		IF fbFaultInjector.Status.xBusy THEN
			iTakeSlot := 1;
			iPutSlot := 1;
			IF fbFaultInjector.xWrongOperation THEN
				eActualOperation := E_MAGAZINE_OPERATION.NONE;
			ELSIF fbFaultInjector.xNoFreeSlot THEN
				eActualOperation := E_MAGAZINE_OPERATION.PUT;
			ELSE
				eActualOperation := E_MAGAZINE_OPERATION.TAKE;
			END_IF;
			Diag.eState := E_MAGAZINE_STATE.CHOOSE;
		ELSIF xFinishedLatched OR xFinishedCondition THEN
			Diag.eState := E_MAGAZINE_STATE.DISABLED;
		// Активный автоматический цикл сначала должен передать владение второму
		// магазину. До этого сохраняем xEnabled + xDisablePending, иначе менеджер
		// остаётся владельцем уже выключенного магазина и не может продолжить груз.
		ELSIF xDisableRequest
		AND NOT xRobotInMagazineContext THEN
			Diag.eState := E_MAGAZINE_STATE.DISABLED;
		ELSIF xGlobalError THEN
			Error.dwErrorActive := Error.dwErrorActive OR ERR_GLOBAL_STOP;
			Diag.eState := E_MAGAZINE_STATE.ERROR;
		// Автоматический владелец держит xExecute до завершения операции. Если
		// команда пришла раньше включения магазина, фронт был бы поглощён в
		// DISABLED; в IDLE принимаем также активный уровень запроса.
		ELSIF (rtExecute.Q OR xExecuteRequest) AND xMechanismReady THEN
			IF xManualCommand THEN
				CASE stHmiCommand.eSetPoint OF
					E_POINT_NAME.MAGAZINE_TAKE_DETAIL:
						eActualOperation := E_MAGAZINE_OPERATION.TAKE;
						iTakeSlot := stHmiCommand.iActiveSlot;
					E_POINT_NAME.MAGAZINE_PUT_DETAIL:
						eActualOperation := E_MAGAZINE_OPERATION.PUT;
						iPutSlot := stHmiCommand.iActiveSlot;
					E_POINT_NAME.MAGAZINE_CHANGE_DETAIL:
						// CHANGE требует двух слотов и запускается через ST_MAGAZINE_COMMAND.
						eActualOperation := E_MAGAZINE_OPERATION.NONE;
					E_POINT_NAME.MAGAZINE_RETURN_BLANK:
						eActualOperation := E_MAGAZINE_OPERATION.RETURN_BLANK;
						iPutSlot := stHmiCommand.iActiveSlot;
				ELSE
						eActualOperation := E_MAGAZINE_OPERATION.NONE;
				END_CASE;
			ELSE
				eActualOperation := stMagazineCommand.eOperation;
				iTakeSlot := stMagazineCommand.iTakeSlot;
				iPutSlot := stMagazineCommand.iPutSlot;
			END_IF;

			Diag.eState := E_MAGAZINE_STATE.CHOOSE;
		END_IF;

	E_MAGAZINE_STATE.CHOOSE:
		xTakeSlotValid := (iTakeSlot >= 1) AND (iTakeSlot <= iActiveSlotCount);
		xPutSlotValid := (iPutSlot >= 1) AND (iPutSlot <= iActiveSlotCount);
		xChangeTakeFirst := (eActualOperation = E_MAGAZINE_OPERATION.CHANGE)
			AND (iTakeSlot = iPutSlot);
		xTakeSlotHasBlank := FALSE;
		xPutSlotEmpty := FALSE;

		IF xTakeSlotValid THEN
		xTakeSlotHasBlank := stInventory.aSlots[iTakeSlot].xInPosition
			AND (stInventory.aSlots[iTakeSlot].eDetailType = E_DETAIL_TYPE.BLANK)
			AND (stInventory.aSlots[iTakeSlot].uiProductType >= UINT#1)
			AND (stInventory.aSlots[iTakeSlot].uiProductType <= uiTypeCount);
		END_IF;

	IF xPutSlotValid THEN
		xPutSlotEmpty := NOT stInventory.aSlots[iPutSlot].xInPosition;
	END_IF;
	xPutProductTypeValid := TRUE;
	IF (eActualOperation = E_MAGAZINE_OPERATION.PUT)
	OR (eActualOperation = E_MAGAZINE_OPERATION.CHANGE) THEN
		xPutProductTypeValid := (stRobotStatus.uiDetailPayloadType >= UINT#1)
			AND (stRobotStatus.uiDetailPayloadType <= uiTypeCount);
	ELSIF eActualOperation = E_MAGAZINE_OPERATION.RETURN_BLANK THEN
		xPutProductTypeValid := (stRobotStatus.uiBlankPayloadType >= UINT#1)
			AND (stRobotStatus.uiBlankPayloadType <= uiTypeCount);
	END_IF;

		IF fbFaultInjector.xGeometry
		OR (iActiveSlotCount = 0) THEN
			Error.dwErrorActive := Error.dwErrorActive OR ERR_GEOMETRY;
			Diag.eState := E_MAGAZINE_STATE.ERROR;

		ELSIF fbFaultInjector.xWrongOperation
		OR (eActualOperation = E_MAGAZINE_OPERATION.NONE) THEN
			Error.dwErrorActive := Error.dwErrorActive OR ERR_WRONG_OPERATION;
			Diag.eState := E_MAGAZINE_STATE.ERROR;

		ELSIF fbFaultInjector.xNoBlank THEN
			Error.dwErrorActive := Error.dwErrorActive OR ERR_NO_BLANK;
			Diag.eState := E_MAGAZINE_STATE.ERROR;

		ELSIF fbFaultInjector.xNoFreeSlot THEN
			Error.dwErrorActive := Error.dwErrorActive OR ERR_NO_FREE_SLOT;
			Diag.eState := E_MAGAZINE_STATE.ERROR;

		ELSIF fbFaultInjector.xInvalidSlot THEN
			Error.dwErrorActive := Error.dwErrorActive OR ERR_INVALID_SLOT;
			Diag.eState := E_MAGAZINE_STATE.ERROR;

		ELSIF fbFaultInjector.xSlotContent THEN
			Error.dwErrorActive := Error.dwErrorActive OR ERR_SLOT_CONTENT;
			Diag.eState := E_MAGAZINE_STATE.ERROR;

		ELSIF ((eActualOperation = E_MAGAZINE_OPERATION.TAKE)
			OR (eActualOperation = E_MAGAZINE_OPERATION.CHANGE))
		AND NOT xTakeSlotValid THEN
			Error.dwErrorActive := Error.dwErrorActive OR ERR_NO_BLANK OR ERR_INVALID_SLOT;
			Diag.eState := E_MAGAZINE_STATE.ERROR;

		ELSIF ((eActualOperation = E_MAGAZINE_OPERATION.PUT)
			OR (eActualOperation = E_MAGAZINE_OPERATION.CHANGE)
			OR (eActualOperation = E_MAGAZINE_OPERATION.RETURN_BLANK))
		AND NOT xPutSlotValid THEN
			Error.dwErrorActive := Error.dwErrorActive OR ERR_NO_FREE_SLOT OR ERR_INVALID_SLOT;
			Diag.eState := E_MAGAZINE_STATE.ERROR;

		ELSIF ((eActualOperation = E_MAGAZINE_OPERATION.TAKE)
			OR (eActualOperation = E_MAGAZINE_OPERATION.CHANGE))
		AND NOT xTakeSlotHasBlank THEN
			Error.dwErrorActive := Error.dwErrorActive OR ERR_SLOT_CONTENT;
			Diag.eState := E_MAGAZINE_STATE.ERROR;

		ELSIF ((eActualOperation = E_MAGAZINE_OPERATION.PUT)
			OR (eActualOperation = E_MAGAZINE_OPERATION.CHANGE)
			OR (eActualOperation = E_MAGAZINE_OPERATION.RETURN_BLANK))
		AND NOT xPutSlotEmpty
		AND NOT (xChangeTakeFirst AND xTakeSlotHasBlank) THEN
			Error.dwErrorActive := Error.dwErrorActive OR ERR_SLOT_CONTENT;
			Diag.eState := E_MAGAZINE_STATE.ERROR;

		ELSIF ((eActualOperation = E_MAGAZINE_OPERATION.PUT)
			OR (eActualOperation = E_MAGAZINE_OPERATION.CHANGE)
			OR (eActualOperation = E_MAGAZINE_OPERATION.RETURN_BLANK))
		AND NOT xPutProductTypeValid THEN
			Error.dwErrorActive := Error.dwErrorActive OR ERR_SLOT_CONTENT;
			Diag.eState := E_MAGAZINE_STATE.ERROR;

		ELSIF (eActualOperation = E_MAGAZINE_OPERATION.TAKE)
		AND (stRobotStatus.xBlankAvailable OR stRobotStatus.xDetailAvailable) THEN
			Error.dwErrorActive := Error.dwErrorActive OR ERR_WRONG_OPERATION;
			Diag.eState := E_MAGAZINE_STATE.ERROR;

		ELSIF (eActualOperation = E_MAGAZINE_OPERATION.CHANGE)
		AND (NOT stRobotStatus.xGripper1Open
			OR stRobotStatus.xBlankAvailable) THEN
			Error.dwErrorActive := Error.dwErrorActive OR ERR_WRONG_OPERATION;
			Diag.eState := E_MAGAZINE_STATE.ERROR;

		ELSIF ((eActualOperation = E_MAGAZINE_OPERATION.PUT)
			OR (eActualOperation = E_MAGAZINE_OPERATION.CHANGE))
		AND NOT stRobotStatus.xDetailAvailable THEN
			Error.dwErrorActive := Error.dwErrorActive OR ERR_WRONG_OPERATION;
			Diag.eState := E_MAGAZINE_STATE.ERROR;

		ELSIF (eActualOperation = E_MAGAZINE_OPERATION.RETURN_BLANK)
		AND (NOT stRobotStatus.xBlankAvailable
			OR stRobotStatus.xDetailAvailable) THEN
			Error.dwErrorActive := Error.dwErrorActive OR ERR_WRONG_OPERATION;
			Diag.eState := E_MAGAZINE_STATE.ERROR;

		ELSE
			uiPutProductType := UINT#0;
			IF (eActualOperation = E_MAGAZINE_OPERATION.PUT)
			OR (eActualOperation = E_MAGAZINE_OPERATION.CHANGE) THEN
				uiPutProductType := stRobotStatus.uiDetailPayloadType;
			ELSIF eActualOperation = E_MAGAZINE_OPERATION.RETURN_BLANK THEN
				uiPutProductType := stRobotStatus.uiBlankPayloadType;
			END_IF;
			xInventoryCommitted := FALSE;
			xTakeSlotCommitted := FALSE;
			xPutSlotCommitted := FALSE;
			xOperationSequenceComplete := FALSE;
			uiStep := 0;
			Diag.eState := E_MAGAZINE_STATE.PREPARE_STEP;
		END_IF;

	E_MAGAZINE_STATE.PREPARE_STEP:
		xRobotCommandStarted := FALSE;
		stActiveRobotCommand.xExecute := FALSE;
		stActiveRobotCommand.xStop := FALSE;
		stActiveRobotCommand.xReset := xResetRequest;
		stActiveRobotCommand.eAction := E_ROBOT_ACTION.NONE;
		stActiveRobotCommand.eSetPoint := E_POINT_NAME.NONE;

		CASE eActualOperation OF
			E_MAGAZINE_OPERATION.TAKE:
				iActiveSlot := iTakeSlot;
			E_MAGAZINE_OPERATION.PUT,
			E_MAGAZINE_OPERATION.RETURN_BLANK:
				iActiveSlot := iPutSlot;
			E_MAGAZINE_OPERATION.CHANGE:
				IF uiStep <= UINT#5 THEN
					iActiveSlot := iPutSlot;
				ELSE
					iActiveSlot := iTakeSlot;
				END_IF;
		ELSE
			iActiveSlot := SINT#0;
		END_CASE;
		stActiveRobotCommand.iActiveSlot := iActiveSlot;
		stActiveRobotCommand.uiMagazineId := uiMagazineId;

		CASE eActualOperation OF
				E_MAGAZINE_OPERATION.TAKE:
					CASE uiStep OF
						0:
							IF stRobotStatus.xRotatedToDetail THEN
								Diag.eState := E_MAGAZINE_STATE.NEXT;
							ELSE
								stActiveRobotCommand.eAction := E_ROBOT_ACTION.ROTATE_TO_DETAIL;
							END_IF;
						1:
							stActiveRobotCommand.eAction := E_ROBOT_ACTION.MOVE_TO_POINT;
							stActiveRobotCommand.eSetPoint := E_POINT_NAME.MAGAZINE_SAFE;
						2:
							stActiveRobotCommand.eAction := E_ROBOT_ACTION.MOVE_TO_POINT;
							stActiveRobotCommand.eSetPoint := E_POINT_NAME.MAGAZINE_IN_SLOT;
						3: stActiveRobotCommand.eAction := E_ROBOT_ACTION.CLAMP_1;
						4:
							stActiveRobotCommand.eAction := E_ROBOT_ACTION.MOVE_TO_POINT;
							stActiveRobotCommand.eSetPoint := E_POINT_NAME.MAGAZINE_SAFE;
					ELSE
						xOperationSequenceComplete := TRUE;
						Diag.eState := E_MAGAZINE_STATE.DONE;
					END_CASE;

				E_MAGAZINE_OPERATION.PUT:
					CASE uiStep OF
						0:
							IF stRobotStatus.xRotatedToBlank THEN
								Diag.eState := E_MAGAZINE_STATE.NEXT;
							ELSE
								stActiveRobotCommand.eAction := E_ROBOT_ACTION.ROTATE_TO_BLANK;
							END_IF;
						1:
							stActiveRobotCommand.eAction := E_ROBOT_ACTION.MOVE_TO_POINT;
							stActiveRobotCommand.eSetPoint := E_POINT_NAME.MAGAZINE_SAFE;
						2:
							stActiveRobotCommand.eAction := E_ROBOT_ACTION.MOVE_TO_POINT;
							stActiveRobotCommand.eSetPoint := E_POINT_NAME.MAGAZINE_IN_SLOT;
						3: stActiveRobotCommand.eAction := E_ROBOT_ACTION.UNCLAMP_2;
						4:
							stActiveRobotCommand.eAction := E_ROBOT_ACTION.MOVE_TO_POINT;
							stActiveRobotCommand.eSetPoint := E_POINT_NAME.MAGAZINE_SAFE;
					ELSE
						xOperationSequenceComplete := TRUE;
						Diag.eState := E_MAGAZINE_STATE.DONE;
					END_CASE;

				E_MAGAZINE_OPERATION.CHANGE:
					CASE uiStep OF
						0:
							IF (xChangeTakeFirst AND stRobotStatus.xRotatedToDetail)
							OR (NOT xChangeTakeFirst AND stRobotStatus.xRotatedToBlank) THEN
								Diag.eState := E_MAGAZINE_STATE.NEXT;
							ELSIF xChangeTakeFirst THEN
								stActiveRobotCommand.eAction := E_ROBOT_ACTION.ROTATE_TO_DETAIL;
							ELSE
								stActiveRobotCommand.eAction := E_ROBOT_ACTION.ROTATE_TO_BLANK;
							END_IF;
						1:
							stActiveRobotCommand.eAction := E_ROBOT_ACTION.MOVE_TO_POINT;
							stActiveRobotCommand.eSetPoint := E_POINT_NAME.MAGAZINE_SAFE;
						2:
							stActiveRobotCommand.eAction := E_ROBOT_ACTION.MOVE_TO_POINT;
							stActiveRobotCommand.eSetPoint := E_POINT_NAME.MAGAZINE_IN_SLOT;
						3:
							IF xChangeTakeFirst THEN
								stActiveRobotCommand.eAction := E_ROBOT_ACTION.CLAMP_1;
							ELSE
								stActiveRobotCommand.eAction := E_ROBOT_ACTION.UNCLAMP_2;
							END_IF;
						4:
							stActiveRobotCommand.eAction := E_ROBOT_ACTION.MOVE_TO_POINT;
							stActiveRobotCommand.eSetPoint := E_POINT_NAME.MAGAZINE_CHANGE;
						5:
							IF (xChangeTakeFirst AND stRobotStatus.xRotatedToBlank)
							OR (NOT xChangeTakeFirst AND stRobotStatus.xRotatedToDetail) THEN
								Diag.eState := E_MAGAZINE_STATE.NEXT;
							ELSIF xChangeTakeFirst THEN
								stActiveRobotCommand.eAction := E_ROBOT_ACTION.ROTATE_TO_BLANK;
							ELSE
								stActiveRobotCommand.eAction := E_ROBOT_ACTION.ROTATE_TO_DETAIL;
							END_IF;
						6:
							stActiveRobotCommand.eAction := E_ROBOT_ACTION.MOVE_TO_POINT;
							stActiveRobotCommand.eSetPoint := E_POINT_NAME.MAGAZINE_CHANGE;
						7:
							stActiveRobotCommand.eAction := E_ROBOT_ACTION.MOVE_TO_POINT;
							stActiveRobotCommand.eSetPoint := E_POINT_NAME.MAGAZINE_IN_SLOT;
						8:
							IF xChangeTakeFirst THEN
								stActiveRobotCommand.eAction := E_ROBOT_ACTION.UNCLAMP_2;
							ELSE
								stActiveRobotCommand.eAction := E_ROBOT_ACTION.CLAMP_1;
							END_IF;
						9:
							stActiveRobotCommand.eAction := E_ROBOT_ACTION.MOVE_TO_POINT;
							stActiveRobotCommand.eSetPoint := E_POINT_NAME.MAGAZINE_SAFE;
					ELSE
						xOperationSequenceComplete := TRUE;
						Diag.eState := E_MAGAZINE_STATE.DONE;
					END_CASE;

				E_MAGAZINE_OPERATION.RETURN_BLANK:
					CASE uiStep OF
						0:
							IF stRobotStatus.xRotatedToDetail THEN
								Diag.eState := E_MAGAZINE_STATE.NEXT;
							ELSE
								stActiveRobotCommand.eAction := E_ROBOT_ACTION.ROTATE_TO_DETAIL;
							END_IF;
						1:
							stActiveRobotCommand.eAction := E_ROBOT_ACTION.MOVE_TO_POINT;
							stActiveRobotCommand.eSetPoint := E_POINT_NAME.MAGAZINE_SAFE;
						2:
							stActiveRobotCommand.eAction := E_ROBOT_ACTION.MOVE_TO_POINT;
							stActiveRobotCommand.eSetPoint := E_POINT_NAME.MAGAZINE_IN_SLOT;
						3: stActiveRobotCommand.eAction := E_ROBOT_ACTION.UNCLAMP_1;
						4:
							stActiveRobotCommand.eAction := E_ROBOT_ACTION.MOVE_TO_POINT;
							stActiveRobotCommand.eSetPoint := E_POINT_NAME.MAGAZINE_SAFE;
					ELSE
						xOperationSequenceComplete := TRUE;
						Diag.eState := E_MAGAZINE_STATE.DONE;
					END_CASE;
		END_CASE;

		IF Diag.eState = E_MAGAZINE_STATE.PREPARE_STEP THEN
			Diag.eState := E_MAGAZINE_STATE.ROBOT_COMMAND;
		END_IF;

	E_MAGAZINE_STATE.ROBOT_COMMAND:
		Command := stActiveRobotCommand;
		Command.xExecute := TRUE;
		IF stRobotStatus.xBusy THEN
			xRobotCommandStarted := TRUE;
		END_IF;

		IF xStopRequest OR xGlobalError THEN
			Command.xStop := stRobotStatus.xBusy;
			Error.dwErrorActive := Error.dwErrorActive OR ERR_GLOBAL_STOP;
			Diag.eState := E_MAGAZINE_STATE.ERROR;

		ELSIF stRobotStatus.xError THEN
			Error.dwErrorActive := Error.dwErrorActive OR ERR_ROBOT;
			Diag.eState := E_MAGAZINE_STATE.ERROR;

		ELSIF xRobotCommandStarted AND stRobotStatus.xDone THEN
			// Матрица меняется в момент подтверждённого физического переноса,
			// а не после отхода робота и завершения всей составной операции.
			CASE eActualOperation OF
				E_MAGAZINE_OPERATION.TAKE:
					IF (uiStep = UINT#3) AND NOT xTakeSlotCommitted THEN
						stInventory.aSlots[iTakeSlot].xInPosition := FALSE;
						stInventory.aSlots[iTakeSlot].eDetailType := E_DETAIL_TYPE.NONE;
						stInventory.aSlots[iTakeSlot].uiProductType := UINT#0;
						xTakeSlotCommitted := TRUE;
					END_IF;

				E_MAGAZINE_OPERATION.PUT:
					IF (uiStep = UINT#3) AND NOT xPutSlotCommitted THEN
						stInventory.aSlots[iPutSlot].xInPosition := TRUE;
						stInventory.aSlots[iPutSlot].eDetailType := E_DETAIL_TYPE.DETAIL;
						stInventory.aSlots[iPutSlot].uiProductType := uiPutProductType;
						udiProducedPartsTotal := udiProducedPartsTotal + UDINT#1;
						xPutSlotCommitted := TRUE;
					END_IF;

				E_MAGAZINE_OPERATION.CHANGE:
					IF (((uiStep = UINT#3) AND NOT xChangeTakeFirst)
						OR ((uiStep = UINT#8) AND xChangeTakeFirst))
					AND NOT xPutSlotCommitted THEN
						stInventory.aSlots[iPutSlot].xInPosition := TRUE;
						stInventory.aSlots[iPutSlot].eDetailType := E_DETAIL_TYPE.DETAIL;
						stInventory.aSlots[iPutSlot].uiProductType := uiPutProductType;
						udiProducedPartsTotal := udiProducedPartsTotal + UDINT#1;
						xPutSlotCommitted := TRUE;
					ELSIF (((uiStep = UINT#8) AND NOT xChangeTakeFirst)
						OR ((uiStep = UINT#3) AND xChangeTakeFirst))
					AND NOT xTakeSlotCommitted THEN
						stInventory.aSlots[iTakeSlot].xInPosition := FALSE;
						stInventory.aSlots[iTakeSlot].eDetailType := E_DETAIL_TYPE.NONE;
						stInventory.aSlots[iTakeSlot].uiProductType := UINT#0;
						xTakeSlotCommitted := TRUE;
					END_IF;

				E_MAGAZINE_OPERATION.RETURN_BLANK:
					IF (uiStep = UINT#3) AND NOT xPutSlotCommitted THEN
						xFinishedLatched := FALSE;
						xFinishedCondition := FALSE;
						stInventory.aSlots[iPutSlot].xInPosition := TRUE;
						stInventory.aSlots[iPutSlot].eDetailType := E_DETAIL_TYPE.BLANK;
						stInventory.aSlots[iPutSlot].uiProductType := uiPutProductType;
						xPutSlotCommitted := TRUE;
					END_IF;
			END_CASE;
			Diag.eState := E_MAGAZINE_STATE.RELEASE_ROBOT_COMMAND;
		END_IF;

	E_MAGAZINE_STATE.RELEASE_ROBOT_COMMAND:
		IF stRobotStatus.xError THEN
			Error.dwErrorActive := Error.dwErrorActive OR ERR_ROBOT;
			Diag.eState := E_MAGAZINE_STATE.ERROR;
		ELSIF NOT stRobotStatus.xBusy AND NOT stRobotStatus.xDone THEN
			Diag.eState := E_MAGAZINE_STATE.NEXT;
		END_IF;

	E_MAGAZINE_STATE.NEXT:
		uiStep := uiStep + 1;
		Diag.eState := E_MAGAZINE_STATE.PREPARE_STEP;

	E_MAGAZINE_STATE.DONE:
		// Страховочная фиксация нужна только если конечный DONE получен без
		// промежуточного обновления. В штатном ходе слоты уже изменены захватами.
		IF xOperationSequenceComplete
		AND NOT xStopRequest
		AND NOT xGlobalError
		AND NOT xInventoryCommitted THEN
			CASE eActualOperation OF
				E_MAGAZINE_OPERATION.TAKE:
					IF NOT xTakeSlotCommitted THEN
						stInventory.aSlots[iTakeSlot].xInPosition := FALSE;
						stInventory.aSlots[iTakeSlot].eDetailType := E_DETAIL_TYPE.NONE;
						stInventory.aSlots[iTakeSlot].uiProductType := UINT#0;
						xTakeSlotCommitted := TRUE;
					END_IF;
				E_MAGAZINE_OPERATION.PUT:
					IF NOT xPutSlotCommitted THEN
						stInventory.aSlots[iPutSlot].xInPosition := TRUE;
						stInventory.aSlots[iPutSlot].eDetailType := E_DETAIL_TYPE.DETAIL;
						stInventory.aSlots[iPutSlot].uiProductType := uiPutProductType;
						udiProducedPartsTotal := udiProducedPartsTotal + UDINT#1;
						xPutSlotCommitted := TRUE;
					END_IF;
				E_MAGAZINE_OPERATION.CHANGE:
					// Для обмена в одном слоте сначала отражаем изъятие. Уже
					// подтверждённую укладку нельзя затереть страховочной фиксацией.
					IF NOT xTakeSlotCommitted THEN
						IF NOT xChangeTakeFirst OR NOT xPutSlotCommitted THEN
							stInventory.aSlots[iTakeSlot].xInPosition := FALSE;
							stInventory.aSlots[iTakeSlot].eDetailType := E_DETAIL_TYPE.NONE;
							stInventory.aSlots[iTakeSlot].uiProductType := UINT#0;
						END_IF;
						xTakeSlotCommitted := TRUE;
					END_IF;
					IF NOT xPutSlotCommitted THEN
						stInventory.aSlots[iPutSlot].xInPosition := TRUE;
						stInventory.aSlots[iPutSlot].eDetailType := E_DETAIL_TYPE.DETAIL;
						stInventory.aSlots[iPutSlot].uiProductType := uiPutProductType;
						udiProducedPartsTotal := udiProducedPartsTotal + UDINT#1;
						xPutSlotCommitted := TRUE;
					END_IF;
				E_MAGAZINE_OPERATION.RETURN_BLANK:
					IF NOT xPutSlotCommitted THEN
						xFinishedLatched := FALSE;
						xFinishedCondition := FALSE;
						stInventory.aSlots[iPutSlot].xInPosition := TRUE;
						stInventory.aSlots[iPutSlot].eDetailType := E_DETAIL_TYPE.BLANK;
						stInventory.aSlots[iPutSlot].uiProductType := uiPutProductType;
						xPutSlotCommitted := TRUE;
					END_IF;
			END_CASE;
			xInventoryCommitted := TRUE;
		END_IF;
		IF NOT xExecuteRequest THEN
			eActualOperation := E_MAGAZINE_OPERATION.NONE;
			IF xDisableRequest
			AND NOT xRobotInMagazineContext THEN
				Diag.eState := E_MAGAZINE_STATE.DISABLED;
			ELSE
				Diag.eState := E_MAGAZINE_STATE.IDLE;
			END_IF;
		END_IF;

	E_MAGAZINE_STATE.ERROR:
		IF xResetRequest
		AND NOT xIoManual
		AND NOT xExecuteRequest
		AND NOT xStopRequest
		AND NOT FaultStatus.xBusy
		AND NOT xGlobalError
		AND xRobotResetDependencyReady THEN
			Error.dwErrorLast := Error.dwErrorActive;
			Error.dwErrorActive := DWORD#0;
			eActualOperation := E_MAGAZINE_OPERATION.NONE;
			Diag.eState := E_MAGAZINE_STATE.DISABLED;
		END_IF;
END_CASE;

// Класс реакции не размазывается по CASE. Первичная причина остаётся в своей
// маске, а контекст конкретного магазина хранится до принятого сброса.
IF (Diag.eState = E_MAGAZINE_STATE.ERROR)
AND NOT xFaultContextCaptured THEN
	xRobotInMagazineAtFault := xRobotInMagazineContext;
	xFaultContextCaptured := TRUE;
ELSIF Diag.eState <> E_MAGAZINE_STATE.ERROR THEN
	xRobotInMagazineAtFault := FALSE;
	xFaultContextCaptured := FALSE;
END_IF;

xRobotStopRequired := NOT xGlobalError
	AND (
		((Error.dwErrorActive AND ERR_ROBOT) <> DWORD#0)
		OR (((Error.dwErrorActive AND MASK_EQUIPMENT_ERROR) <> DWORD#0)
			AND xRobotInMagazineAtFault)
	);

// Физический Stop нужен только занятому роботу. При неподвижном роботе внутри
// магазина FB_ROBOT получит зависимую ошибку без пустой команды остановки.
IF (Diag.eState = E_MAGAZINE_STATE.ERROR)
AND xRobotStopRequired
AND stRobotStatus.xBusy THEN
	Command := stActiveRobotCommand;
	Command.xExecute := TRUE;
	Command.xStop := TRUE;
END_IF;

// ERROR технологически отключает магазин немедленно, но причина остаётся
// защёлкнутой до разрешённого Reset.
Status.xEnabled := (Diag.eState <> E_MAGAZINE_STATE.DISABLED)
	AND (Diag.eState <> E_MAGAZINE_STATE.ERROR);
Status.xDisablePending := xDisableRequest AND Status.xEnabled;
Status.xPowerAllowed := Status.xEnabled OR Status.xEnableSequenceAllowed;
Status.xFillAllowed := (iActiveSlotCount > SINT#0) AND Status.xEditAllowed;
Status.xClearAllowed := Status.xEditAllowed;
Status.xReady := xMechanismReady AND  (Diag.eState = E_MAGAZINE_STATE.IDLE)
	AND xRobotCanWorkWithMagazine
	AND (Error.dwErrorActive = DWORD#0);
Status.xBusy := (Diag.eState <> E_MAGAZINE_STATE.DISABLED)
	AND (Diag.eState <> E_MAGAZINE_STATE.IDLE)
	AND (Diag.eState <> E_MAGAZINE_STATE.DONE)
	AND (Diag.eState <> E_MAGAZINE_STATE.ERROR);
Status.xDone := Diag.eState = E_MAGAZINE_STATE.DONE;
Status.xError := Diag.eState = E_MAGAZINE_STATE.ERROR;
Status.xRobotStopRequired := xRobotStopRequired;
Status.udiProducedPartsTotal := udiProducedPartsTotal;
Status.uiMagazineId := uiMagazineId;
Status.eGrantedOperation := eGrantedOperation;
Status.eActualOperation := eActualOperation;
Status.iSelectedBlank := iTakeSlot;
Status.iSelectedFreeSlot := iPutSlot;
// Разовая доработка палеты завершена: чужой груз/станок не возвращает её
// в планирование. Защёлку снимает только смена банка или правка его содержимого.
xFinishedLatched := xFinishedLatched OR (xFinishedCondition AND NOT Status.xBusy);
Status.xFinished := xFinishedLatched;
Error.dwAlarmActive := Error.dwErrorActive;

IF Error.dwErrorActive <> DWORD#0 THEN
	Error.dwErrorLast := Error.dwErrorActive;
END_IF;

Error.stErrorActive := UpdateErrorView(dwError := Error.dwErrorActive);
Error.stErrorLast := UpdateErrorView(dwError := Error.dwErrorLast);
FaultStatus.xResetAllowed := Status.xError
	AND NOT xIoManual
	AND NOT FaultStatus.xBusy
	AND NOT xExecuteRequest
	AND NOT xStopRequest
	AND NOT xGlobalError
	AND xRobotResetDependencyReady;

// Сводка публикуется владельцем содержимого после всех изменений слотов.
UpdateTypeStatus(stMagazineInventory := stInventory);

METHOD FindBlank : SINT
VAR_INPUT
	iSlotCount : SINT; // Число слотов, участвующих в поиске
END_VAR
VAR_IN_OUT
	stDetail : ARRAY [1..GVL_CELL_SETTINGS.NumberDetail] OF ST_DETAIL; // Содержимое слотов магазина
END_VAR
VAR
	i : SINT; // Индекс проверяемого слота
END_VAR
FindBlank := 0;

FOR i:= 1 TO iSlotCount DO
	IF stDetail[i].xInPosition = TRUE AND stDetail[i].eDetailType =  E_DETAIL_TYPE.BLANK THEN
		FindBlank := i;
		EXIT;
	END_IF
END_FOR
END_METHOD

METHOD UpdateErrorView : ST_MAGAZINE_ERROR
VAR_INPUT
	dwError : DWORD; // Битовая маска для расшифровки
END_VAR
VAR
	stError : ST_MAGAZINE_ERROR; // Представление ошибок отдельными флагами
END_VAR
stError.WRONG_OPERATION := (dwError AND ERR_WRONG_OPERATION) <> DWORD#0;
stError.NO_BLANK := (dwError AND ERR_NO_BLANK) <> DWORD#0;
stError.NO_FREE_SLOT := (dwError AND ERR_NO_FREE_SLOT) <> DWORD#0;
stError.INVALID_SLOT := (dwError AND ERR_INVALID_SLOT) <> DWORD#0;
stError.SLOT_CONTENT := (dwError AND ERR_SLOT_CONTENT) <> DWORD#0;
stError.ROBOT_ERROR := (dwError AND ERR_ROBOT) <> DWORD#0;
stError.GLOBAL_STOP := (dwError AND ERR_GLOBAL_STOP) <> DWORD#0;
stError.GEOMETRY_ERROR := (dwError AND ERR_GEOMETRY) <> DWORD#0;

UpdateErrorView := stError;
END_METHOD

METHOD FindFreeSlot : SINT
VAR_INPUT
	iSlotCount : SINT; // Число слотов, участвующих в поиске
END_VAR
VAR_IN_OUT
	stDetail : ARRAY [1..GVL_CELL_SETTINGS.NumberDetail] OF ST_DETAIL; // Содержимое слотов магазина
END_VAR
VAR
	i : SINT; // Индекс проверяемого слота
END_VAR
FindFreeSlot := 0;

FOR i:= 1 TO iSlotCount DO
	IF stDetail[i].xInPosition = FALSE THEN
		FindFreeSlot := i;
		EXIT;
	END_IF
END_FOR
END_METHOD

METHOD PRIVATE UpdateTypeStatus
VAR_IN_OUT
	stMagazineInventory : ST_MAGAZINE_INVENTORY;
END_VAR
VAR
	uiType : UINT; // Тип секции, 1..3
	uiSlot : UINT; // Проверяемый слот
	iSlot  : SINT; // Индекс массива содержимого
END_VAR
FOR uiType := UINT#1 TO UINT#3 DO
	Status.stTypeStatus.aiBlankSlot[uiType] := SINT#0;
	Status.stTypeStatus.aiFreeSlot[uiType] := SINT#0;
	Status.stTypeStatus.auiBlankCount[uiType] := UINT#0;
	Status.stTypeStatus.auiDetailCount[uiType] := UINT#0;
	Status.stTypeStatus.auiFreeCount[uiType] := UINT#0;
END_FOR;

IF (iActiveSlotCount > SINT#0)
AND (uiTypeCount >= UINT#1)
AND (uiTypeCount <= UINT#3) THEN
	FOR uiSlot := UINT#1 TO SINT_TO_UINT(iActiveSlotCount) DO
		iSlot := UINT_TO_SINT(uiSlot);
		IF NOT stMagazineInventory.aSlots[iSlot].xInPosition THEN
			// Пустой слот универсален: тип 0
			// означает отсутствие изделия, а не запрет укладки конкретного типа.
			FOR uiType := UINT#1 TO uiTypeCount DO
				Status.stTypeStatus.auiFreeCount[uiType] :=
					Status.stTypeStatus.auiFreeCount[uiType] + UINT#1;
				IF Status.stTypeStatus.aiFreeSlot[uiType] = SINT#0 THEN
					Status.stTypeStatus.aiFreeSlot[uiType] := iSlot;
				END_IF;
			END_FOR;
		ELSE
			uiType := stMagazineInventory.aSlots[iSlot].uiProductType;
			IF (uiType >= UINT#1) AND (uiType <= uiTypeCount)
			AND (stMagazineInventory.aSlots[iSlot].eDetailType = E_DETAIL_TYPE.BLANK) THEN
				Status.stTypeStatus.auiBlankCount[uiType] :=
					Status.stTypeStatus.auiBlankCount[uiType] + UINT#1;
				IF Status.stTypeStatus.aiBlankSlot[uiType] = SINT#0 THEN
					Status.stTypeStatus.aiBlankSlot[uiType] := iSlot;
				END_IF;
			ELSIF (uiType >= UINT#1) AND (uiType <= uiTypeCount)
			AND (stMagazineInventory.aSlots[iSlot].eDetailType = E_DETAIL_TYPE.DETAIL) THEN
				Status.stTypeStatus.auiDetailCount[uiType] :=
					Status.stTypeStatus.auiDetailCount[uiType] + UINT#1;
			END_IF;
		END_IF;
	END_FOR;
END_IF;
END_METHOD

END_FUNCTION_BLOCK

// Device/Application/FB/FB_FAULT_INJECTOR/FB_MAGAZINE_FAULT_INJECTOR
FUNCTION_BLOCK FB_MAGAZINE_FAULT_INJECTOR
VAR_INPUT
	Request       : ST_MAGAZINE_FAULT_REQUEST; // Запросы конкретных ошибок магазина
	xOwnerAllowed : BOOL; // Безопасные условия, рассчитанные FB_MAGAZINE
	xComplete     : BOOL; // Штатная ошибка уже сформирована владельцем
END_VAR
VAR_OUTPUT
	xWrongOperation : BOOL;
	xNoBlank        : BOOL;
	xNoFreeSlot     : BOOL;
	xInvalidSlot    : BOOL;
	xSlotContent    : BOOL;
	xGeometry       : BOOL;
	Status          : ST_FAULT_INJECTION_STATUS; // Состояние источника для HMI
END_VAR
VAR
	rtWrongOperation : R_TRIG;
	rtNoBlank        : R_TRIG;
	rtNoFreeSlot     : R_TRIG;
	rtInvalidSlot    : R_TRIG;
	rtSlotContent    : R_TRIG;
	rtGeometry       : R_TRIG;
	xRequestPulse    : BOOL;
END_VAR

rtWrongOperation(CLK := Request.xWrongOperation);
rtNoBlank(CLK := Request.xNoBlank);
rtNoFreeSlot(CLK := Request.xNoFreeSlot);
rtInvalidSlot(CLK := Request.xInvalidSlot);
rtSlotContent(CLK := Request.xSlotContent);
rtGeometry(CLK := Request.xGeometry);

xRequestPulse := rtWrongOperation.Q
	OR rtNoBlank.Q
	OR rtNoFreeSlot.Q
	OR rtInvalidSlot.Q
	OR rtSlotContent.Q
	OR rtGeometry.Q;

Status.xRejected := FALSE;
Status.xAllowed := Request.xEnabled AND xOwnerAllowed;

IF xComplete THEN
	xWrongOperation := FALSE;
	xNoBlank := FALSE;
	xNoFreeSlot := FALSE;
	xInvalidSlot := FALSE;
	xSlotContent := FALSE;
	xGeometry := FALSE;
END_IF;

IF xRequestPulse THEN
	IF Status.xAllowed THEN
		xWrongOperation := rtWrongOperation.Q;
		xNoBlank := rtNoBlank.Q;
		xNoFreeSlot := rtNoFreeSlot.Q;
		xInvalidSlot := rtInvalidSlot.Q;
		xSlotContent := rtSlotContent.Q;
		xGeometry := rtGeometry.Q;
	ELSE
		Status.xRejected := TRUE;
		Status.udiRejectSequence := Status.udiRejectSequence + UDINT#1;
		IF Status.udiRejectSequence = UDINT#0 THEN
			Status.udiRejectSequence := UDINT#1;
		END_IF;
	END_IF;
END_IF;

Status.xActive := xWrongOperation
	OR xNoBlank
	OR xNoFreeSlot
	OR xInvalidSlot
	OR xSlotContent
	OR xGeometry;
Status.xBusy := Status.xActive;
Status.xResetAllowed := FALSE;

END_FUNCTION_BLOCK

// Device/Application/FB/FB_ROBOT_MODBUS
{attribute 'no_assign'}
FUNCTION_BLOCK FB_ROBOT_MODBUS
VAR_INPUT
	xEnable          : BOOL; // Применён режим MODBUS_TCP
	xReconnect       : BOOL; // Настройки изменены, выполнить reconnect
	Config           : ST_ROBOT_MODBUS_CONFIG;
	Command          : ST_ROBOT_COMMAND; // Семантическая команда FB_ROBOT
END_VAR
VAR_OUTPUT
	Status           : ST_ROBOT_MODBUS_STATUS;
END_VAR
VAR_IN_OUT
	auiWriteRegisters : ARRAY [0..8] OF UINT; // Документные адреса 1001..1009
	auiReadRegisters  : ARRAY [0..16] OF UINT; // Документные адреса 1101..1117
END_VAR
VAR
	{attribute 'no_assign'}
	fbClient       : ModbusFB.ClientTCP;
	fbRead         : ModbusFB.ClientRequestReadHoldingRegisters;
	fbWrite        : ModbusFB.ClientRequestWriteMultipleRegisters;
	eState         : E_ROBOT_MODBUS_CLIENT_STATE := E_ROBOT_MODBUS_CLIENT_STATE.DISABLED;
	xConnect       : BOOL;
	xReadExecute   : BOOL;
	xWriteExecute  : BOOL;
	xStatusFresh   : BOOL;
	xCommandArmed  : BOOL;
	xCommandActive : BOOL;
	xWritePending  : BOOL;
	xHeartbeatChanged : BOOL;
	xHeartbeatSeen : BOOL;
	xPlcHeartbeatDue : BOOL;
	xStopPending   : BOOL;
	xResetPending  : BOOL;
	xResetInProgress : BOOL;
	xResetWriteDone : BOOL; // FC16 с Reset=1 подтверждена сервером
	tonResetAttempt : TON;
	xControlClearPending : BOOL;
	rtStop         : R_TRIG;
	rtReset        : R_TRIG;
	rtReconnect    : R_TRIG;
	tonPoll        : TON;
	tonPlcHeartbeat: TON;
	tonRobotHeartbeat : TON;
	tonCommunicationGrace : TON;
	tonCommandTimeout : TON;
	tonReconnect   : TON;
	uiCommandSeq   : UINT;
	uiActiveSeq    : UINT;
	uiDecodedRobotHeartbeat : UINT; // Heartbeat из последнего завершённого FC03
	uiPositionXHigh : UINT; // Координаты из того же завершённого FC03-снимка
	uiPositionXLow  : UINT;
	uiPositionYHigh : UINT;
	uiPositionYLow  : UINT;
	uiPositionZHigh : UINT;
	uiPositionZLow  : UINT;
	uiPlcHeartbeat : UINT;
	uiLastRobotHeartbeat : UINT;
	uiCommandCode  : UINT;
	uiRegisterIndex : UINT;
	dwPositionRaw  : DWORD;
	diPositionRaw  : DINT;
	udiReplyTimeoutUs : UDINT;
END_VAR
VAR CONSTANT
	COMMAND_START_ITEM : UINT := UINT#1000; // Документный 1001
	STATUS_START_ITEM  : UINT := UINT#1100; // Документный 1101
	COMMAND_QUANTITY   : UINT := UINT#9;
	STATUS_QUANTITY    : UINT := UINT#17;
	PROTOCOL_VERSION   : UINT := UINT#3;
	RESET_ATTEMPT_TIMEOUT : TIME := T#10S; // Полная попытка: запись, feedback, снятие
	STATUS_CONTROLLER_ON  : UINT := UINT#16#0001;
	STATUS_AUTOMATIC_MODE : UINT := UINT#16#0002;
	STATUS_REMOTE_ENABLED : UINT := UINT#16#0004;
	STATUS_DRIVES_ENABLED : UINT := UINT#16#0008;
	STATUS_HOMED          : UINT := UINT#16#0010;
	STATUS_EMERGENCY_STOP : UINT := UINT#16#0020;
	STATUS_ROBOT_ALARM    : UINT := UINT#16#0040;
	STATUS_ROBOT_READY    : UINT := UINT#16#0080;
	STATUS_POSITION_VALID : UINT := UINT#16#0100;
	STATUS_SIMULATOR_ACTIVE : UINT := UINT#16#0200;
END_VAR

Status.xConfigValid := (Config.aIpAddress[0] > BYTE#0)
	AND (Config.aIpAddress[0] < BYTE#224)
	AND (Config.uiPort > UINT#0)
	AND (Config.uiUnitId <= UINT#255)
	AND (Config.tResponseTimeout >= T#50MS)
	AND (Config.tPollInterval >= T#10MS)
	AND (Config.tHeartbeatTimeout >= T#500MS)
	AND (Config.tCommandTimeout >= T#1S);

	udiReplyTimeoutUs := TIME_TO_UDINT(Config.tResponseTimeout) * UDINT#1000;
	rtStop(CLK := Command.xStop);
	rtReset(CLK := Command.xReset);
	rtReconnect(CLK := xReconnect);
	IF rtStop.Q THEN
		xStopPending := TRUE;
	END_IF;
	IF rtReset.Q AND NOT xResetInProgress THEN
		xResetPending := TRUE;
		xResetInProgress := TRUE;
		xResetWriteDone := FALSE;
		Status.xResetDone := FALSE;
		Status.xResetFailed := FALSE;
	END_IF;
xReadExecute := FALSE;
xWriteExecute := FALSE;
xHeartbeatChanged := FALSE;

fbClient(
	xConnect := xConnect,
	aIPaddr := Config.aIpAddress,
	uiPort := Config.uiPort,
	tConnnectTimeOut := Config.tHeartbeatTimeout
);

IF NOT xEnable OR NOT Status.xConfigValid THEN
	xConnect := FALSE;
	eState := E_ROBOT_MODBUS_CLIENT_STATE.DISABLED;
	xStatusFresh := FALSE;
	xCommandArmed := FALSE;
	xCommandActive := FALSE;
	xWritePending := FALSE;
	xStopPending := FALSE;
	xResetPending := FALSE;
	xResetInProgress := FALSE;
	xResetWriteDone := FALSE;
	Status.xResetDone := FALSE;
	Status.xResetFailed := FALSE;
	xControlClearPending := FALSE;
	xHeartbeatSeen := FALSE;
	xPlcHeartbeatDue := FALSE;
	uiActiveSeq := UINT#0;
	Status.xConnected := FALSE;
ELSE
	xConnect := TRUE;
	IF rtReconnect.Q THEN
		xConnect := FALSE;
		eState := E_ROBOT_MODBUS_CLIENT_STATE.RECONNECT_WAIT;
		xStatusFresh := FALSE;
		xCommandArmed := FALSE;
		xCommandActive := FALSE;
		xWritePending := FALSE;
		xControlClearPending := FALSE;
		xHeartbeatSeen := FALSE;
		xPlcHeartbeatDue := FALSE;
	END_IF;
END_IF;

CASE eState OF
	E_ROBOT_MODBUS_CLIENT_STATE.DISABLED:
		IF xEnable AND Status.xConfigValid THEN
			xConnect := TRUE;
			eState := E_ROBOT_MODBUS_CLIENT_STATE.CONNECTING;
		END_IF;

	E_ROBOT_MODBUS_CLIENT_STATE.CONNECTING:
		IF fbClient.xConnected THEN
			eState := E_ROBOT_MODBUS_CLIENT_STATE.INITIAL_READ;
		ELSIF fbClient.xError THEN
			Status.udiClientError := TO_UDINT(fbClient.eErrorID);
			xConnect := FALSE;
			eState := E_ROBOT_MODBUS_CLIENT_STATE.RECONNECT_WAIT;
		END_IF;

	E_ROBOT_MODBUS_CLIENT_STATE.INITIAL_READ:
		xReadExecute := TRUE;
		IF fbRead.xDone THEN
			xStatusFresh := TRUE;
			uiCommandSeq := auiReadRegisters[0];
			uiActiveSeq := UINT#0;
			uiPlcHeartbeat := UINT#0;
			uiLastRobotHeartbeat := auiReadRegisters[6];
			xHeartbeatSeen := FALSE;
			FOR uiRegisterIndex := UINT#0 TO UINT#8 DO
				auiWriteRegisters[uiRegisterIndex] := UINT#0;
			END_FOR;
			auiWriteRegisters[7] := uiCommandSeq;
			eState := E_ROBOT_MODBUS_CLIENT_STATE.INITIAL_READ_RELEASE;
		ELSIF fbRead.xError THEN
			Status.udiReadError := TO_UDINT(fbRead.eErrorID);
			xConnect := FALSE;
			eState := E_ROBOT_MODBUS_CLIENT_STATE.RECONNECT_WAIT;
		END_IF;

	E_ROBOT_MODBUS_CLIENT_STATE.INITIAL_READ_RELEASE:
		IF NOT fbRead.xBusy THEN
			eState := E_ROBOT_MODBUS_CLIENT_STATE.CLEAR_COMMAND;
		END_IF;

	E_ROBOT_MODBUS_CLIENT_STATE.CLEAR_COMMAND:
		xWriteExecute := TRUE;
		IF fbWrite.xDone THEN
			eState := E_ROBOT_MODBUS_CLIENT_STATE.CLEAR_COMMAND_RELEASE;
		ELSIF fbWrite.xError THEN
			Status.udiWriteError := TO_UDINT(fbWrite.eErrorID);
			xConnect := FALSE;
			eState := E_ROBOT_MODBUS_CLIENT_STATE.RECONNECT_WAIT;
		END_IF;

	E_ROBOT_MODBUS_CLIENT_STATE.CLEAR_COMMAND_RELEASE:
		IF NOT fbWrite.xBusy THEN
			xCommandArmed := NOT Command.xExecute;
			xCommandActive := FALSE;
			eState := E_ROBOT_MODBUS_CLIENT_STATE.READY;
		END_IF;

	E_ROBOT_MODBUS_CLIENT_STATE.READY:
		IF NOT fbClient.xConnected OR fbClient.xError THEN
			Status.udiClientError := TO_UDINT(fbClient.eErrorID);
			xConnect := FALSE;
			eState := E_ROBOT_MODBUS_CLIENT_STATE.RECONNECT_WAIT;
		ELSIF xStopPending THEN
			// Stop отменяет текущую попытку сброса; он не может быть проглочен Reset.
			IF xResetInProgress THEN Status.xResetFailed := TRUE; END_IF;
			xResetInProgress := FALSE;
			xResetWriteDone := FALSE;
			// Stop always preempts Reset and normal commands.
			// Execute снимается сразу: после принятого CommandSeq это не отменяет
			// команду, зато позволяет роботу выйти из DONE/ERROR/STOPPED в IDLE.
			// Без этого уже завершённая дискретная команда навечно удерживала
			// Execute=1, а xControlClearPending ждал недостижимый IDLE.
			auiWriteRegisters[0] := UINT#0;
			auiWriteRegisters[1] := UINT#0;
			auiWriteRegisters[2] := UINT#1;
			auiWriteRegisters[3] := UINT#0;
			auiWriteRegisters[4] := UINT#0;
			auiWriteRegisters[5] := UINT#0;
			auiWriteRegisters[6] := UINT#0;
			xStopPending := FALSE;
			xResetPending := FALSE;
			xControlClearPending := TRUE;
			xWritePending := TRUE;
		ELSIF xResetPending THEN
			// Reset обязан прервать незавершённую очистку Stop. Иначе
			// xControlClearPending имеет приоритет и защёлкнутый Reset никогда
			// не попадает в регистр 1004.
			auiWriteRegisters[0] := UINT#0;
			auiWriteRegisters[1] := UINT#0;
			auiWriteRegisters[2] := UINT#0;
			auiWriteRegisters[3] := UINT#1;
			auiWriteRegisters[4] := UINT#0;
			auiWriteRegisters[5] := UINT#0;
			auiWriteRegisters[6] := UINT#0;
			xCommandActive := FALSE;
			uiActiveSeq := UINT#0;
			xCommandArmed := FALSE;
			xResetPending := FALSE;
			xControlClearPending := TRUE;
			xWritePending := TRUE;
		ELSIF xControlClearPending THEN
			// Stop удерживается до STOPPED/IDLE, Reset — до снятия аварии. Так
			// импульс не потеряется между более медленными циклами программы робота.
			IF ((auiWriteRegisters[2] = UINT#1)
				AND ((Status.uiExecutionState = TO_UINT(E_ROBOT_MODBUS_EXECUTION_STATE.STOPPED))
					OR (Status.uiExecutionState = TO_UINT(E_ROBOT_MODBUS_EXECUTION_STATE.IDLE))))
			OR ((auiWriteRegisters[3] = UINT#1)
				AND xResetWriteDone
				AND NOT Status.xRobotAlarm
				AND (Status.uiExecutionState =
					TO_UINT(E_ROBOT_MODBUS_EXECUTION_STATE.IDLE))) THEN
				auiWriteRegisters[2] := UINT#0;
				auiWriteRegisters[3] := UINT#0;
				xCommandActive := FALSE;
				uiActiveSeq := UINT#0;
				// Верхний FB удерживает Execute до появления Busy. Поэтому после
				// подтверждённой очистки принимаем уже удерживаемую новую команду,
				// а не требуем ещё одного фронта от HMI.
				xCommandArmed := TRUE;
				xControlClearPending := FALSE;
				xWritePending := TRUE;
			END_IF;
		ELSIF Command.xExecute AND xCommandArmed AND NOT xCommandActive THEN
			uiCommandCode := UINT#0;
			CASE Command.eAction OF
				E_ROBOT_ACTION.MOVE_TO_POINT:
					CASE Command.eSetPoint OF
						E_POINT_NAME.MACHINE_1_ABOVE: uiCommandCode := UINT#10;
						E_POINT_NAME.MACHINE_1_INSIDE: uiCommandCode := UINT#11;
						E_POINT_NAME.MACHINE_1_CHUCK_APROACH: uiCommandCode := UINT#12;
						E_POINT_NAME.MACHINE_1_CHUCK_POSITION: uiCommandCode := UINT#13;
						E_POINT_NAME.MACHINE_2_ABOVE: uiCommandCode := UINT#14;
						E_POINT_NAME.MACHINE_2_INSIDE: uiCommandCode := UINT#15;
						E_POINT_NAME.MACHINE_2_CHUCK_APROACH: uiCommandCode := UINT#16;
						E_POINT_NAME.MACHINE_2_CHUCK_POSITION: uiCommandCode := UINT#17;
						E_POINT_NAME.MACHINE_3_ABOVE: uiCommandCode := UINT#18;
						E_POINT_NAME.MACHINE_3_INSIDE: uiCommandCode := UINT#19;
						E_POINT_NAME.MACHINE_3_CHUCK_APROACH: uiCommandCode := UINT#20;
						E_POINT_NAME.MACHINE_3_CHUCK_POSITION: uiCommandCode := UINT#21;
						E_POINT_NAME.HOME_SAFETY: uiCommandCode := UINT#22;
						E_POINT_NAME.MAGAZINE_SAFE: uiCommandCode := UINT#23;
						E_POINT_NAME.MAGAZINE_CHANGE: uiCommandCode := UINT#24;
						E_POINT_NAME.MAGAZINE_IN_SLOT: uiCommandCode := UINT#25;
					END_CASE;
				E_ROBOT_ACTION.UNCLAMP_1: uiCommandCode := UINT#2;
				E_ROBOT_ACTION.CLAMP_1: uiCommandCode := UINT#3;
				E_ROBOT_ACTION.UNCLAMP_2: uiCommandCode := UINT#4;
				E_ROBOT_ACTION.CLAMP_2: uiCommandCode := UINT#5;
				E_ROBOT_ACTION.ROTATE_TO_BLANK: uiCommandCode := UINT#6;
				E_ROBOT_ACTION.ROTATE_TO_DETAIL: uiCommandCode := UINT#7;
			END_CASE;

			IF uiCommandCode > UINT#0 THEN
				uiCommandSeq := uiCommandSeq + UINT#1;
				IF uiCommandSeq = UINT#0 THEN
					uiCommandSeq := UINT#1;
				END_IF;
				uiActiveSeq := uiCommandSeq;
				auiWriteRegisters[0] := uiCommandCode;
				auiWriteRegisters[1] := UINT#1;
				auiWriteRegisters[2] := UINT#0;
				auiWriteRegisters[3] := UINT#0;
				auiWriteRegisters[4] := SINT_TO_UINT(Command.iActiveSlot);
				auiWriteRegisters[5] := Command.uiMagazineId;
				auiWriteRegisters[6] := UINT#0;
				auiWriteRegisters[7] := uiCommandSeq;
				xCommandActive := TRUE;
				xCommandArmed := FALSE;
				xWritePending := TRUE;
			END_IF;
		ELSIF NOT Command.xExecute AND xCommandActive THEN
			auiWriteRegisters[0] := UINT#0;
			auiWriteRegisters[1] := UINT#0;
			auiWriteRegisters[2] := UINT#0;
			auiWriteRegisters[3] := UINT#0;
			auiWriteRegisters[4] := UINT#0;
			auiWriteRegisters[5] := UINT#0;
			auiWriteRegisters[6] := UINT#0;
			xCommandActive := FALSE;
			// CommandSeq в регистре сохраняется как последний использованный номер,
			// но завершённая транзакция больше не имеет права публиковать Done.
			// Повтор после Reset всегда получит новый ненулевой sequence.
			uiActiveSeq := UINT#0;
			xCommandArmed := TRUE;
			xWritePending := TRUE;
		ELSIF NOT Command.xExecute THEN
			xCommandArmed := TRUE;
		END_IF;

		IF xPlcHeartbeatDue THEN
			uiPlcHeartbeat := uiPlcHeartbeat + UINT#1;
			auiWriteRegisters[8] := uiPlcHeartbeat;
			xPlcHeartbeatDue := FALSE;
			xWritePending := TRUE;
		END_IF;

		IF xWritePending THEN
			eState := E_ROBOT_MODBUS_CLIENT_STATE.WRITE_COMMAND;
		ELSIF tonPoll.Q THEN
			eState := E_ROBOT_MODBUS_CLIENT_STATE.READ_STATUS;
		END_IF;

	E_ROBOT_MODBUS_CLIENT_STATE.WRITE_COMMAND:
		xWriteExecute := TRUE;
		IF fbWrite.xDone THEN
			IF xResetInProgress THEN
				IF auiWriteRegisters[3] = UINT#1 THEN
					xResetWriteDone := TRUE;
				ELSIF xResetWriteDone AND NOT xControlClearPending THEN
					// Успех только после FC03 без аварии/с IDLE и последующей
					// подтверждённой записи Reset=0. Один локальный скан не Ack.
					xResetInProgress := FALSE;
					Status.xResetDone := TRUE;
				END_IF;
			END_IF;
			xWritePending := FALSE;
			eState := E_ROBOT_MODBUS_CLIENT_STATE.WRITE_COMMAND_RELEASE;
		ELSIF fbWrite.xError THEN
			Status.udiWriteError := TO_UDINT(fbWrite.eErrorID);
			xConnect := FALSE;
			eState := E_ROBOT_MODBUS_CLIENT_STATE.RECONNECT_WAIT;
		END_IF;

	E_ROBOT_MODBUS_CLIENT_STATE.WRITE_COMMAND_RELEASE:
		IF NOT fbWrite.xBusy THEN
			eState := E_ROBOT_MODBUS_CLIENT_STATE.READ_STATUS;
		END_IF;

	E_ROBOT_MODBUS_CLIENT_STATE.READ_STATUS:
		xReadExecute := TRUE;
		IF fbRead.xDone THEN
			xStatusFresh := TRUE;
			eState := E_ROBOT_MODBUS_CLIENT_STATE.READ_STATUS_RELEASE;
		ELSIF fbRead.xError THEN
			Status.udiReadError := TO_UDINT(fbRead.eErrorID);
			xConnect := FALSE;
			eState := E_ROBOT_MODBUS_CLIENT_STATE.RECONNECT_WAIT;
		END_IF;

	E_ROBOT_MODBUS_CLIENT_STATE.READ_STATUS_RELEASE:
		IF NOT fbRead.xBusy THEN
			eState := E_ROBOT_MODBUS_CLIENT_STATE.READY;
		END_IF;

	E_ROBOT_MODBUS_CLIENT_STATE.RECONNECT_WAIT:
		xConnect := FALSE;
		xStatusFresh := FALSE;
		IF tonReconnect.Q THEN
			xConnect := TRUE;
			eState := E_ROBOT_MODBUS_CLIENT_STATE.CONNECTING;
		END_IF;
END_CASE;

tonResetAttempt(IN := xResetInProgress, PT := RESET_ATTEMPT_TIMEOUT);
IF xResetInProgress
AND ((eState = E_ROBOT_MODBUS_CLIENT_STATE.RECONNECT_WAIT)
	OR rtReconnect.Q OR tonResetAttempt.Q OR NOT Command.xReset) THEN
	// Не повторяем неоднозначную запись после обрыва. Reconnect сначала
	// прочитает состояние и очистит блок; новый Reset требует нового фронта.
	xResetInProgress := FALSE;
	xResetPending := FALSE;
	xResetWriteDone := FALSE;
	Status.xResetDone := FALSE;
	Status.xResetFailed := TRUE;
	xConnect := FALSE;
	xStatusFresh := FALSE;
	eState := E_ROBOT_MODBUS_CLIENT_STATE.RECONNECT_WAIT;
END_IF;
IF eState = E_ROBOT_MODBUS_CLIENT_STATE.RECONNECT_WAIT THEN
	xReadExecute := FALSE;
	xWriteExecute := FALSE;
	xControlClearPending := FALSE;
	xWritePending := FALSE;
	xCommandArmed := FALSE;
END_IF;
Status.xResetBusy := xResetInProgress;

fbRead(
	xExecute := xReadExecute,
	udiTimeOut := udiReplyTimeoutUs,
	rClient := fbClient,
	uiUnitId := Config.uiUnitId,
	udiReplyTimeout := udiReplyTimeoutUs,
	uiMaxRetries := UINT#1,
	uiStartItem := STATUS_START_ITEM,
	uiQuantity := STATUS_QUANTITY,
	pData := ADR(auiReadRegisters)
);
fbWrite(
	xExecute := xWriteExecute,
	udiTimeOut := udiReplyTimeoutUs,
	rClient := fbClient,
	uiUnitId := Config.uiUnitId,
	udiReplyTimeout := udiReplyTimeoutUs,
	uiMaxRetries := UINT#1,
	uiStartItem := COMMAND_START_ITEM,
	uiQuantity := COMMAND_QUANTITY,
	pData := ADR(auiWriteRegisters)
);

// FC03 может завершиться внутри вызова fbRead. Декодирование выполняется после
// вызова, чтобы технологический Status и сырые диагностические регистры всегда
// относились к одному и тому же снимку опроса.
IF fbRead.xDone THEN
	Status.uiAckSeq := auiReadRegisters[0];
	Status.uiExecutionState := auiReadRegisters[1];
	Status.uiResultCode := auiReadRegisters[2];
	Status.uiActiveCommand := auiReadRegisters[3];
	Status.uiCurrentPoint := auiReadRegisters[4];
	Status.uiGripperStatus := auiReadRegisters[5];
	Status.uiRobotHeartbeat := auiReadRegisters[6];
	Status.uiStatusWord := auiReadRegisters[7];
	Status.uiAlarmCode := auiReadRegisters[8];
	Status.uiOperationPhase := auiReadRegisters[15];
	Status.uiProtocolVersion := auiReadRegisters[16];
	uiDecodedRobotHeartbeat := auiReadRegisters[6];
	uiPositionXHigh := auiReadRegisters[9];
	uiPositionXLow := auiReadRegisters[10];
	uiPositionYHigh := auiReadRegisters[11];
	uiPositionYLow := auiReadRegisters[12];
	uiPositionZHigh := auiReadRegisters[13];
	uiPositionZLow := auiReadRegisters[14];
END_IF;

tonPoll(IN := eState = E_ROBOT_MODBUS_CLIENT_STATE.READY, PT := Config.tPollInterval);
// Heartbeat timer is independent of request states. The due latch prevents a pulse
// from being lost while FC03/FC16 is busy.
tonPlcHeartbeat(
	IN := xEnable AND fbClient.xConnected AND NOT tonPlcHeartbeat.Q,
	PT := T#100MS
);
IF tonPlcHeartbeat.Q THEN
	xPlcHeartbeatDue := TRUE;
END_IF;
tonReconnect(IN := eState = E_ROBOT_MODBUS_CLIENT_STATE.RECONNECT_WAIT, PT := T#1S);

Status.xConnected := fbClient.xConnected AND xConnect;
Status.xStatusFresh := xStatusFresh;

IF uiDecodedRobotHeartbeat <> uiLastRobotHeartbeat THEN
	uiLastRobotHeartbeat := uiDecodedRobotHeartbeat;
	xHeartbeatChanged := TRUE;
	xHeartbeatSeen := TRUE;
END_IF;
tonRobotHeartbeat(
	IN := xEnable AND xStatusFresh AND NOT xHeartbeatChanged,
	PT := Config.tHeartbeatTimeout
);
Status.xCommunicationAlive := Status.xConnected
	AND xStatusFresh
	AND xHeartbeatSeen
	AND NOT tonRobotHeartbeat.Q
	AND (Status.uiProtocolVersion = PROTOCOL_VERSION);
tonCommunicationGrace(
	IN := xEnable AND Status.xConfigValid AND NOT Status.xCommunicationAlive,
	PT := Config.tHeartbeatTimeout
);

Status.xControllerOn := (Status.uiStatusWord AND STATUS_CONTROLLER_ON) <> UINT#0;
Status.xAutomaticMode := (Status.uiStatusWord AND STATUS_AUTOMATIC_MODE) <> UINT#0;
Status.xRemoteEnabled := (Status.uiStatusWord AND STATUS_REMOTE_ENABLED) <> UINT#0;
Status.xDrivesEnabled := (Status.uiStatusWord AND STATUS_DRIVES_ENABLED) <> UINT#0;
Status.xHomed := (Status.uiStatusWord AND STATUS_HOMED) <> UINT#0;
Status.xEmergencyStop := (Status.uiStatusWord AND STATUS_EMERGENCY_STOP) <> UINT#0;
Status.xRobotAlarm := ((Status.uiStatusWord AND STATUS_ROBOT_ALARM) <> UINT#0)
	OR (Status.uiAlarmCode <> UINT#0);
Status.xPositionValid := (Status.uiStatusWord AND STATUS_POSITION_VALID) <> UINT#0;
Status.xSimulatorActive := (Status.uiStatusWord AND STATUS_SIMULATOR_ACTIVE) <> UINT#0;
Status.xReady := Status.xCommunicationAlive
	AND Status.xControllerOn
	AND Status.xAutomaticMode
	AND Status.xRemoteEnabled
	AND Status.xDrivesEnabled
	AND Status.xHomed
	AND Status.xPositionValid
	AND NOT Status.xEmergencyStop
	AND NOT Status.xRobotAlarm
	AND ((Status.uiStatusWord AND STATUS_ROBOT_READY) <> UINT#0);

Status.xDone := (uiActiveSeq <> UINT#0)
	AND xCommandActive
	AND (Status.uiAckSeq = uiActiveSeq)
	AND (Status.uiExecutionState = TO_UINT(E_ROBOT_MODBUS_EXECUTION_STATE.DONE))
	AND (Status.uiResultCode = UINT#0);
// Busy означает активную PLC-транзакцию, включая ожидание AckSeq. Благодаря
// этому FB_ROBOT обязательно увидит запуск новой команды до её terminal state.
Status.xBusy := (uiActiveSeq <> UINT#0)
	AND xCommandActive
	AND NOT Status.xDone
	AND NOT ((Status.uiAckSeq = uiActiveSeq)
		AND ((Status.uiExecutionState = TO_UINT(E_ROBOT_MODBUS_EXECUTION_STATE.ERROR))
			OR (Status.uiExecutionState = TO_UINT(E_ROBOT_MODBUS_EXECUTION_STATE.STOPPED))
			OR ((Status.uiExecutionState = TO_UINT(E_ROBOT_MODBUS_EXECUTION_STATE.DONE))
				AND (Status.uiResultCode <> UINT#0))));
tonCommandTimeout(
	IN := xCommandActive AND NOT Status.xDone,
	PT := Config.tCommandTimeout
);
Status.xCommandTimeout := tonCommandTimeout.Q;
Status.xError := tonCommunicationGrace.Q
	OR Status.xResetFailed
	OR Status.xRobotAlarm
	OR Status.xCommandTimeout
	OR ((uiActiveSeq <> UINT#0)
		AND (Status.uiAckSeq = uiActiveSeq)
		AND ((Status.uiExecutionState = TO_UINT(E_ROBOT_MODBUS_EXECUTION_STATE.ERROR))
			OR ((Status.uiExecutionState = TO_UINT(E_ROBOT_MODBUS_EXECUTION_STATE.DONE))
				AND (Status.uiResultCode <> UINT#0))));

dwPositionRaw := SHL(UINT_TO_DWORD(uiPositionXHigh), 16)
	OR UINT_TO_DWORD(uiPositionXLow);
diPositionRaw := DWORD_TO_DINT(dwPositionRaw);
Status.lrActualX := DINT_TO_LREAL(diPositionRaw) / LREAL#10.0;
dwPositionRaw := SHL(UINT_TO_DWORD(uiPositionYHigh), 16)
	OR UINT_TO_DWORD(uiPositionYLow);
diPositionRaw := DWORD_TO_DINT(dwPositionRaw);
Status.lrActualY := DINT_TO_LREAL(diPositionRaw) / LREAL#10.0;
dwPositionRaw := SHL(UINT_TO_DWORD(uiPositionZHigh), 16)
	OR UINT_TO_DWORD(uiPositionZLow);
diPositionRaw := DWORD_TO_DINT(dwPositionRaw);
Status.lrActualZ := DINT_TO_LREAL(diPositionRaw) / LREAL#10.0;

END_FUNCTION_BLOCK

// Device/Application/FB/FB_GRIPPER_SIMULATION
FUNCTION_BLOCK FB_GRIPPER_SIMULATION
VAR_INPUT
	xUsePhysicalFeedback : BOOL; // NORMAL SoftMotion: подтверждать реальные датчики
	xPhysicalIoReady : BOOL;
	PhysicalFeedback : ST_GRIPPER_STATUS;
	tPhysicalActionTimeout : TIME := T#10S;
	xTestInitialize : BOOL;
	auiTestContent : ARRAY [1..2] OF UINT;
	uiTestOrientation : UINT;
	xSimulationAccelerationEnable : BOOL; // Разрешить ускорение таймеров только в симуляции
	uiSimulationTimeFactor : UINT := 1; // Коэффициент виртуального времени 1..100
	Command : ST_GRIPPER_COMMAND; // Команда управления захватом
	FaultRequest : ST_GRIPPER_FAULT_REQUEST; // Единый контракт диагностической инъекции

    tGripper1OpenTime  : TIME := T#500MS; // Время открытия первого захвата
    tGripper1CloseTime : TIME := T#500MS; // Время закрытия первого захвата
    tGripper2OpenTime  : TIME := T#500MS; // Время открытия второго захвата
    tGripper2CloseTime : TIME := T#500MS; // Время закрытия второго захвата
    tRotateTime        : TIME := T#700MS; // Время смены рабочего захвата
END_VAR
VAR_OUTPUT
	Status : ST_GRIPPER_STATUS; // Рабочие статусы захвата
	Diag   : ST_GRIPPER_DIAG; // Состояние автомата и активное действие
	Error  : ST_GRIPPER_ERRORS; // Активные и последние ошибки
	FaultStatus : ST_FAULT_INJECTION_STATUS; // Состояние источника для HMI
END_VAR
VAR
	uiEffectiveTimeFactor : UINT;
	udiActionTime : UDINT;
	fbFaultInjector : FB_GRIPPER_FAULT_INJECTOR; // Изоляция тестовых источников от автомата
	eState        : E_GRIPPER_STATE := E_GRIPPER_STATE.IDLE; // Текущее состояние автомата захвата
    eActiveAction : E_ROBOT_ACTION := E_ROBOT_ACTION.NONE; // Выполняемое действие захвата

    tonAction      : TON; // Таймер выполнения действия
    xActionFault   : BOOL; // Неисправность, относящаяся к текущему действию
	xActionValid   : BOOL; // Получено допустимое действие захвата
    xActionRequired: BOOL; // Для действия требуется физическое переключение
    tActionTime    : TIME; // Нормативное время текущего действия
	xActionConfirmed : BOOL;
	xPhysicalGlobalFault : BOOL;
	xPhysicalGripper1Fault : BOOL;
	xPhysicalGripper2Fault : BOOL;
	xPhysicalRotationFault : BOOL;
    xInitialized   : BOOL; // Начальные состояния установлены
	rtReset         : R_TRIG; // Фронт команды сброса захвата
END_VAR
VAR CONSTANT 
	ERR_GRIPPER_1   : DWORD := DWORD#16#0000_0001; // Ошибка первого захвата
    ERR_GRIPPER_2   : DWORD := DWORD#16#0000_0002; // Ошибка второго захвата
    ERR_GRIP_ROTATE : DWORD := DWORD#16#0000_0004; // Ошибка механизма поворота
    ERR_GRIP_ACTION : DWORD := DWORD#16#0000_0008; // Недопустимое действие захвата
    ERR_GRIP_GLOBAL : DWORD := DWORD#16#0000_0010; // Общая ошибка захвата
	WRN_RESET_EXECUTE_ACTIVE : UINT := 1; // Команда захвата ещё активна
	WRN_RESET_GLOBAL_FAULT   : UINT := 2; // Общая неисправность ещё активна
	WRN_RESET_GRIPPER_1_FAULT: UINT := 3; // Неисправность первого захвата ещё активна
	WRN_RESET_GRIPPER_2_FAULT: UINT := 4; // Неисправность второго захвата ещё активна
	WRN_RESET_ROTATION_FAULT : UINT := 5; // Неисправность поворота ещё активна
END_VAR

uiEffectiveTimeFactor := uiSimulationTimeFactor;
IF NOT xSimulationAccelerationEnable THEN
	uiEffectiveTimeFactor := UINT#1;
ELSIF uiEffectiveTimeFactor < UINT#1 THEN
	uiEffectiveTimeFactor := UINT#1;
ELSIF uiEffectiveTimeFactor > UINT#100 THEN
	uiEffectiveTimeFactor := UINT#100;
END_IF;

IF NOT xInitialized THEN
    Status.xGripper1Open := TRUE;
    Status.xGripper1Closed := FALSE;

    Status.xGripper2Open := TRUE;
    Status.xGripper2Closed := FALSE;

    Status.xRotatedToBlank := TRUE;
    Status.xRotatedToDetail := FALSE;

    xInitialized := TRUE;
END_IF;

IF xTestInitialize THEN
	Status.xGripper1Open := auiTestContent[1] = UINT#0;
	Status.xGripper1Closed := NOT Status.xGripper1Open;
	Status.xGripper2Open := auiTestContent[2] = UINT#0;
	Status.xGripper2Closed := NOT Status.xGripper2Open;
	Status.xRotatedToBlank := uiTestOrientation = UINT#0;
	Status.xRotatedToDetail := NOT Status.xRotatedToBlank;
	eState := E_GRIPPER_STATE.IDLE;
	Error.dwErrorActive := DWORD#0;
END_IF;

// Не создаём подтверждение позиции по прошедшему времени в NORMAL.
IF xUsePhysicalFeedback THEN
	Status.xGripper1Open := PhysicalFeedback.xGripper1Open;
	Status.xGripper1Closed := PhysicalFeedback.xGripper1Closed;
	Status.xGripper2Open := PhysicalFeedback.xGripper2Open;
	Status.xGripper2Closed := PhysicalFeedback.xGripper2Closed;
	Status.xRotatedToBlank := PhysicalFeedback.xRotatedToBlank;
	Status.xRotatedToDetail := PhysicalFeedback.xRotatedToDetail;
END_IF;
xPhysicalGlobalFault := xUsePhysicalFeedback AND NOT xPhysicalIoReady;
xPhysicalGripper1Fault := xUsePhysicalFeedback AND Status.xGripper1Open AND Status.xGripper1Closed;
xPhysicalGripper2Fault := xUsePhysicalFeedback AND Status.xGripper2Open AND Status.xGripper2Closed;
xPhysicalRotationFault := xUsePhysicalFeedback AND Status.xRotatedToBlank AND Status.xRotatedToDetail;

// Ошибочная обратная связь блокирует владельца и до начала действия.
// Используем существующие биты GRIPPER и принятый эффект ROBOT_STOP.
IF xPhysicalGlobalFault THEN
	Error.dwErrorActive := Error.dwErrorActive OR ERR_GRIP_GLOBAL;
	eState := E_GRIPPER_STATE.ERROR;
END_IF;
IF xPhysicalGripper1Fault THEN
	Error.dwErrorActive := Error.dwErrorActive OR ERR_GRIPPER_1;
	eState := E_GRIPPER_STATE.ERROR;
END_IF;
IF xPhysicalGripper2Fault THEN
	Error.dwErrorActive := Error.dwErrorActive OR ERR_GRIPPER_2;
	eState := E_GRIPPER_STATE.ERROR;
END_IF;
IF xPhysicalRotationFault THEN
	Error.dwErrorActive := Error.dwErrorActive OR ERR_GRIP_ROTATE;
	eState := E_GRIPPER_STATE.ERROR;
END_IF;

rtReset(CLK := Command.xReset);

fbFaultInjector(
	Request := FaultRequest,
	eActiveAction := eActiveAction
);
FaultStatus := fbFaultInjector.Status;

IF rtReset.Q
AND (eState = E_GRIPPER_STATE.ERROR) THEN
	IF Command.xExecute THEN
		Diag.stWarning.uiCode := WRN_RESET_EXECUTE_ACTIVE;
	ELSIF fbFaultInjector.xGlobalFault OR xPhysicalGlobalFault THEN
		Diag.stWarning.uiCode := WRN_RESET_GLOBAL_FAULT;
	ELSIF fbFaultInjector.xGripper1Fault OR xPhysicalGripper1Fault THEN
		Diag.stWarning.uiCode := WRN_RESET_GRIPPER_1_FAULT;
	ELSIF fbFaultInjector.xGripper2Fault OR xPhysicalGripper2Fault THEN
		Diag.stWarning.uiCode := WRN_RESET_GRIPPER_2_FAULT;
	ELSIF fbFaultInjector.xRotationFault OR xPhysicalRotationFault THEN
		Diag.stWarning.uiCode := WRN_RESET_ROTATION_FAULT;
	ELSE
		Diag.stWarning.uiCode := UINT#0;
	END_IF;

	IF Diag.stWarning.uiCode <> UINT#0 THEN
		Diag.stWarning.udiSequence := Diag.stWarning.udiSequence + UDINT#1;
		IF Diag.stWarning.udiSequence = UDINT#0 THEN
			Diag.stWarning.udiSequence := UDINT#1;
		END_IF;
	END_IF;
END_IF;


xActionFault := fbFaultInjector.xActionFault;
xActionConfirmed := FALSE;
CASE eActiveAction OF
	E_ROBOT_ACTION.UNCLAMP_1:
		xActionConfirmed := Status.xGripper1Open AND NOT Status.xGripper1Closed;
		xActionFault := xActionFault OR xPhysicalGripper1Fault;
	E_ROBOT_ACTION.CLAMP_1:
		xActionConfirmed := Status.xGripper1Closed AND NOT Status.xGripper1Open;
		xActionFault := xActionFault OR xPhysicalGripper1Fault;
	E_ROBOT_ACTION.UNCLAMP_2:
		xActionConfirmed := Status.xGripper2Open AND NOT Status.xGripper2Closed;
		xActionFault := xActionFault OR xPhysicalGripper2Fault;
	E_ROBOT_ACTION.CLAMP_2:
		xActionConfirmed := Status.xGripper2Closed AND NOT Status.xGripper2Open;
		xActionFault := xActionFault OR xPhysicalGripper2Fault;
	E_ROBOT_ACTION.ROTATE_TO_BLANK:
		xActionConfirmed := Status.xRotatedToBlank AND NOT Status.xRotatedToDetail;
		xActionFault := xActionFault OR xPhysicalRotationFault;
	E_ROBOT_ACTION.ROTATE_TO_DETAIL:
		xActionConfirmed := Status.xRotatedToDetail AND NOT Status.xRotatedToBlank;
		xActionFault := xActionFault OR xPhysicalRotationFault;
END_CASE;
tActionTime := T#0S;

CASE eActiveAction OF
	E_ROBOT_ACTION.UNCLAMP_1:
		tActionTime := tGripper1OpenTime;
	E_ROBOT_ACTION.CLAMP_1:
		tActionTime := tGripper1CloseTime;
	E_ROBOT_ACTION.UNCLAMP_2:
		tActionTime := tGripper2OpenTime;
	E_ROBOT_ACTION.CLAMP_2:
		tActionTime := tGripper2CloseTime;
	E_ROBOT_ACTION.ROTATE_TO_BLANK,
	E_ROBOT_ACTION.ROTATE_TO_DETAIL:
		tActionTime := tRotateTime;

END_CASE;

	udiActionTime := TIME_TO_UDINT(tActionTime) / TO_UDINT(uiEffectiveTimeFactor);
	IF udiActionTime < UDINT#1 THEN
		udiActionTime := UDINT#1;
	END_IF;
	tActionTime := UDINT_TO_TIME(udiActionTime);


IF xUsePhysicalFeedback THEN
	tActionTime := tPhysicalActionTimeout;
END_IF;

tonAction(
    IN := (eState = E_GRIPPER_STATE.EXECUTE)
          AND NOT xActionFault
          AND NOT fbFaultInjector.xGlobalFault AND NOT xPhysicalGlobalFault,
    PT := tActionTime
);


CASE eState OF

    E_GRIPPER_STATE.IDLE:

        Status.xBusy := FALSE;
        Status.xDone := FALSE;
        Status.xError := FALSE;

        IF Command.xExecute THEN
            eActiveAction := Command.eAction;
			xActionValid := TRUE;
			xActionRequired := TRUE;

            CASE Command.eAction OF

				E_ROBOT_ACTION.UNCLAMP_1:
					xActionRequired := NOT (Status.xGripper1Open AND NOT Status.xGripper1Closed);

				E_ROBOT_ACTION.CLAMP_1:
					xActionRequired := NOT (Status.xGripper1Closed AND NOT Status.xGripper1Open);

				E_ROBOT_ACTION.UNCLAMP_2:
					xActionRequired := NOT (Status.xGripper2Open AND NOT Status.xGripper2Closed);

				E_ROBOT_ACTION.CLAMP_2:
					xActionRequired := NOT (Status.xGripper2Closed AND NOT Status.xGripper2Open);

				E_ROBOT_ACTION.ROTATE_TO_BLANK:
					xActionRequired := NOT (Status.xRotatedToBlank AND NOT Status.xRotatedToDetail);

				E_ROBOT_ACTION.ROTATE_TO_DETAIL:
					xActionRequired := NOT (Status.xRotatedToDetail AND NOT Status.xRotatedToBlank);

            ELSE
				xActionValid := FALSE;
                Error.dwErrorActive := Error.dwErrorActive OR ERR_GRIP_ACTION;
                eState := E_GRIPPER_STATE.ERROR;
            END_CASE;

			IF xActionValid THEN
				IF xActionRequired THEN
					eState := E_GRIPPER_STATE.EXECUTE;
				ELSE
					eState := E_GRIPPER_STATE.DONE;
				END_IF;
			END_IF;
        END_IF;


    E_GRIPPER_STATE.EXECUTE:

        Status.xBusy := TRUE;
        Status.xDone := FALSE;

		// Снятие Execute отменяет только незавершённое виртуальное действие и
		// сохраняет последнюю подтверждённую позицию захвата.
		IF NOT Command.xExecute THEN
			Status.xBusy := FALSE;
			eActiveAction := E_ROBOT_ACTION.NONE;
			eState := E_GRIPPER_STATE.IDLE;

		ELSIF fbFaultInjector.xGlobalFault OR xPhysicalGlobalFault THEN
            Error.dwErrorActive := Error.dwErrorActive OR ERR_GRIP_GLOBAL;
            eState := E_GRIPPER_STATE.ERROR;

        ELSIF xActionFault THEN

            CASE eActiveAction OF

                E_ROBOT_ACTION.UNCLAMP_1,
                E_ROBOT_ACTION.CLAMP_1:
                    Error.dwErrorActive := Error.dwErrorActive OR ERR_GRIPPER_1;

                E_ROBOT_ACTION.UNCLAMP_2,
                E_ROBOT_ACTION.CLAMP_2:
                    Error.dwErrorActive := Error.dwErrorActive OR ERR_GRIPPER_2;

                E_ROBOT_ACTION.ROTATE_TO_BLANK,
                E_ROBOT_ACTION.ROTATE_TO_DETAIL:
                    Error.dwErrorActive := Error.dwErrorActive OR ERR_GRIP_ROTATE;

            END_CASE;

            eState := E_GRIPPER_STATE.ERROR;

        ELSIF xUsePhysicalFeedback THEN
			IF xActionConfirmed THEN
				eState := E_GRIPPER_STATE.DONE;
			ELSIF tonAction.Q THEN
				CASE eActiveAction OF
					E_ROBOT_ACTION.UNCLAMP_1, E_ROBOT_ACTION.CLAMP_1:
						Error.dwErrorActive := Error.dwErrorActive OR ERR_GRIPPER_1;
					E_ROBOT_ACTION.UNCLAMP_2, E_ROBOT_ACTION.CLAMP_2:
						Error.dwErrorActive := Error.dwErrorActive OR ERR_GRIPPER_2;
					E_ROBOT_ACTION.ROTATE_TO_BLANK, E_ROBOT_ACTION.ROTATE_TO_DETAIL:
						Error.dwErrorActive := Error.dwErrorActive OR ERR_GRIP_ROTATE;
				END_CASE;
				eState := E_GRIPPER_STATE.ERROR;
			END_IF;

        ELSIF tonAction.Q THEN

            CASE eActiveAction OF

                E_ROBOT_ACTION.UNCLAMP_1:
                    Status.xGripper1Open := TRUE;
                    Status.xGripper1Closed := FALSE;

                E_ROBOT_ACTION.CLAMP_1:
                    Status.xGripper1Open := FALSE;
                    Status.xGripper1Closed := TRUE;

                E_ROBOT_ACTION.UNCLAMP_2:
                    Status.xGripper2Open := TRUE;
                    Status.xGripper2Closed := FALSE;

                E_ROBOT_ACTION.CLAMP_2:
                    Status.xGripper2Open := FALSE;
                    Status.xGripper2Closed := TRUE;

                E_ROBOT_ACTION.ROTATE_TO_BLANK:
                    Status.xRotatedToBlank := TRUE;
                    Status.xRotatedToDetail := FALSE;

                E_ROBOT_ACTION.ROTATE_TO_DETAIL:
                    Status.xRotatedToBlank := FALSE;
                    Status.xRotatedToDetail := TRUE;

            END_CASE;

            eState := E_GRIPPER_STATE.DONE;
        END_IF;


    E_GRIPPER_STATE.DONE:

        Status.xBusy := FALSE;
        Status.xDone := TRUE;

        IF NOT Command.xExecute THEN
            Status.xDone := FALSE;
            eActiveAction := E_ROBOT_ACTION.NONE;
            eState := E_GRIPPER_STATE.IDLE;
        END_IF;


    E_GRIPPER_STATE.ERROR:

        Status.xBusy := FALSE;
        Status.xDone := FALSE;
        Status.xError := TRUE;

        IF Command.xReset
        AND NOT Command.xExecute
        AND NOT fbFaultInjector.xGlobalFault
        AND NOT fbFaultInjector.xGripper1Fault
		AND NOT fbFaultInjector.xGripper2Fault
		AND NOT fbFaultInjector.xRotationFault
		AND NOT xPhysicalGlobalFault
		AND NOT xPhysicalGripper1Fault
		AND NOT xPhysicalGripper2Fault
		AND NOT xPhysicalRotationFault THEN

			Error.dwErrorLast := Error.dwErrorActive;
            Error.dwErrorActive := DWORD#0;
            Status.xError := FALSE;
            eActiveAction := E_ROBOT_ACTION.NONE;
            eState := E_GRIPPER_STATE.IDLE;
        END_IF;

END_CASE;

Diag.eState := eState;
Diag.eActiveAction := eActiveAction;

IF Error.dwErrorActive <> DWORD#0 THEN
	Error.dwErrorLast := Error.dwErrorActive;
END_IF;

Error.stErrorActive := UpdateErrorView(dwError := Error.dwErrorActive);
Error.stErrorLast := UpdateErrorView(dwError := Error.dwErrorLast);
Error.dwAlarmActive := Error.dwErrorActive;
FaultStatus.xResetAllowed := (Error.dwErrorActive <> DWORD#0)
	AND NOT FaultStatus.xActive
	AND NOT xPhysicalGlobalFault
	AND NOT xPhysicalGripper1Fault
	AND NOT xPhysicalGripper2Fault
	AND NOT xPhysicalRotationFault;

METHOD UpdateErrorView : ST_GRIPPER_ERROR
VAR_INPUT
	dwError : DWORD; // Битовая маска для расшифровки
END_VAR
VAR
	stError : ST_GRIPPER_ERROR; // Представление ошибок отдельными флагами
END_VAR
stError.GRIPPER_1_ERROR := (dwError AND ERR_GRIPPER_1) <> DWORD#0;
stError.GRIPPER_2_ERROR := (dwError AND ERR_GRIPPER_2) <> DWORD#0;
stError.ROTATION_ERROR := (dwError AND ERR_GRIP_ROTATE) <> DWORD#0;
stError.ACTION_ERROR := (dwError AND ERR_GRIP_ACTION) <> DWORD#0;
stError.GLOBAL_ERROR := (dwError AND ERR_GRIP_GLOBAL) <> DWORD#0;

UpdateErrorView := stError;
END_METHOD

END_FUNCTION_BLOCK

// Device/Application/FB/FB_FAULT_INJECTOR/FB_GRIPPER_FAULT_INJECTOR
FUNCTION_BLOCK FB_GRIPPER_FAULT_INJECTOR
VAR_INPUT
	Request       : ST_GRIPPER_FAULT_REQUEST; // Поддерживаемые неисправности захвата
	eActiveAction : E_ROBOT_ACTION; // Текущее действие виртуального захвата
END_VAR
VAR_OUTPUT
	xGripper1Fault : BOOL; // Действующая неисправность первого захвата
	xGripper2Fault : BOOL; // Действующая неисправность второго захвата
	xRotationFault : BOOL; // Действующая неисправность поворота
	xGlobalFault   : BOOL; // Действующая общая неисправность
	xActionFault   : BOOL; // Неисправность относится к текущему действию
	Status         : ST_FAULT_INJECTION_STATUS; // Состояние источника для HMI
END_VAR

xGripper1Fault := Request.xEnabled AND Request.xGripper1Fault;
xGripper2Fault := Request.xEnabled AND Request.xGripper2Fault;
xRotationFault := Request.xEnabled AND Request.xRotationFault;
xGlobalFault := Request.xEnabled AND Request.xGlobalFault;

xActionFault := FALSE;
CASE eActiveAction OF
	E_ROBOT_ACTION.UNCLAMP_1,
	E_ROBOT_ACTION.CLAMP_1:
		xActionFault := xGripper1Fault;

	E_ROBOT_ACTION.UNCLAMP_2,
	E_ROBOT_ACTION.CLAMP_2:
		xActionFault := xGripper2Fault;

	E_ROBOT_ACTION.ROTATE_TO_BLANK,
	E_ROBOT_ACTION.ROTATE_TO_DETAIL:
		xActionFault := xRotationFault;
END_CASE;

Status.xAllowed := Request.xEnabled;
Status.xActive := xGripper1Fault
	OR xGripper2Fault
	OR xRotationFault
	OR xGlobalFault;
Status.xBusy := FALSE;
Status.xResetAllowed := NOT Status.xActive;
Status.xRejected := FALSE;

END_FUNCTION_BLOCK

// Device/Application/FB/FB_FAULT_INJECTOR/FB_ROBOT_FAULT_INJECTOR
FUNCTION_BLOCK FB_ROBOT_FAULT_INJECTOR
VAR_INPUT
	Request       : ST_ROBOT_FAULT_REQUEST; // Запросы локальных ошибок робота
	xOwnerAllowed : BOOL; // Безопасные условия, рассчитанные FB_ROBOT
END_VAR
VAR_OUTPUT
	xWrongAction : BOOL; // Одноцикловая недопустимая команда для штатной проверки
	Status       : ST_FAULT_INJECTION_STATUS; // Состояние источника для HMI
END_VAR
VAR
	rtWrongAction : R_TRIG; // Фронт команды HMI
END_VAR

rtWrongAction(CLK := Request.xWrongAction);
xWrongAction := FALSE;
Status.xRejected := FALSE;
Status.xAllowed := Request.xEnabled AND xOwnerAllowed;
Status.xBusy := FALSE;
Status.xResetAllowed := FALSE;

IF rtWrongAction.Q THEN
	IF Status.xAllowed THEN
		xWrongAction := TRUE;
	ELSE
		Status.xRejected := TRUE;
		Status.udiRejectSequence := Status.udiRejectSequence + UDINT#1;
		IF Status.udiRejectSequence = UDINT#0 THEN
			Status.udiRejectSequence := UDINT#1;
		END_IF;
	END_IF;
END_IF;

Status.xActive := xWrongAction;

END_FUNCTION_BLOCK

// Device/Application/FB/FB_MACHINE_SIMULATION
FUNCTION_BLOCK FB_MACHINE_SIMULATION
VAR_INPUT
	xTestInitialize : BOOL;
	uiTestInitialState : UINT;
	xSafetyDoorOpen : BOOL; // Принудительно удерживать операторскую дверь открытой для инъекции
	xSimulationAccelerationEnable : BOOL; // Разрешить ускорение таймеров только в симуляции
	uiSimulationTimeFactor : UINT := 1; // До x250 для автоматических тестов Python-Modbus
    Command : ST_MACHINE_IO_COMMAND; // Команды исполнительным механизмам
	FaultRequest : ST_MACHINE_FAULT_REQUEST; // Единый контракт диагностической инъекции

    tDoorOpenTime   : TIME := T#1S; // Время открытия роботного люка
    tDoorCloseTime  : TIME := T#1S; // Время закрытия роботного люка
    tChuckOpenTime  : TIME := T#1S; // Время разжима патрона
    tChuckCloseTime : TIME := T#1S; // Время зажима патрона
    tCycleTime : TIME := T#47S; // Время цикла обработки
END_VAR

VAR_OUTPUT
    Status : ST_MACHINE_IO_STATUS; // Состояние исполнительных механизмов
	Diag   : ST_MACHINE_SIM_DIAG; // Текущие действия симулятора
	Error  : ST_MACHINE_SIM_ERRORS; // Активные и последние ошибки
END_VAR
VAR CONSTANT
	ERR_MACHINE_ALARM : DWORD := DWORD#16#0000_0001; // Авария станка
	ERR_DOOR_FAULT    : DWORD := DWORD#16#0000_0002; // Ошибка двери
	ERR_CHUCK_FAULT   : DWORD := DWORD#16#0000_0004; // Ошибка патрона
END_VAR

VAR
	uiEffectiveTimeFactor : UINT;
	udiDoorOpenTime : UDINT;
	udiDoorCloseTime : UDINT;
	udiChuckOpenTime : UDINT;
	udiChuckCloseTime : UDINT;
	udiCycleStartTime : UDINT;
	udiCycleTime : UDINT;
	tEffectiveDoorOpenTime : TIME;
	tEffectiveDoorCloseTime : TIME;
	tEffectiveChuckOpenTime : TIME;
	tEffectiveChuckCloseTime : TIME;
	tEffectiveCycleStartTime : TIME;
	tEffectiveCycleTime : TIME;
    rtStartCycle : R_TRIG; // Фронт команды запуска цикла

    tonDoorOpen   : TON; // Таймер открытия двери
    tonDoorClose  : TON; // Таймер закрытия двери
	tonHatchUnlock : TON; // Таймер снятия замка роботного люка
	tonSafetyDoorOpen  : TON; // Таймер открытия операторской двери
	tonSafetyDoorClose : TON; // Таймер закрытия операторской двери
    tonChuckClamp : TON; // Таймер зажима патрона
    tonChuckOpen  : TON; // Таймер разжима патрона
    tonCycleStart : TON; // Таймер подтверждения запуска цикла
    tonCycle      : TON; // Таймер обработки

    xDoorOpening   : BOOL; // Выполняется открытие двери
    xDoorClosing   : BOOL; // Выполняется закрытие двери
	xHatchUnlocking : BOOL; // Выполняется открытие замка
	xSafetyDoorOpening : BOOL; // Выполняется открытие операторской двери
	xSafetyDoorClosing : BOOL; // Выполняется закрытие операторской двери
    xChuckClamping : BOOL; // Выполняется зажим патрона
    xChuckOpening  : BOOL; // Выполняется разжим патрона
    xCycleStarting : BOOL; // Выполняется запуск цикла

    xAlarmLatched : BOOL; // Защёлкнутая авария симулятора
    xInitialized  : BOOL; // Начальные состояния установлены
	xResetRequest : BOOL; // Локальный или переданный станком запрос сброса
END_VAR

uiEffectiveTimeFactor := uiSimulationTimeFactor;
IF NOT xSimulationAccelerationEnable THEN
	uiEffectiveTimeFactor := UINT#1;
ELSIF uiEffectiveTimeFactor < UINT#1 THEN
	uiEffectiveTimeFactor := UINT#1;
ELSIF uiEffectiveTimeFactor > UINT#250 THEN
	uiEffectiveTimeFactor := UINT#250;
END_IF;

udiDoorOpenTime := TIME_TO_UDINT(tDoorOpenTime) / TO_UDINT(uiEffectiveTimeFactor);
udiDoorCloseTime := TIME_TO_UDINT(tDoorCloseTime) / TO_UDINT(uiEffectiveTimeFactor);
udiChuckOpenTime := TIME_TO_UDINT(tChuckOpenTime) / TO_UDINT(uiEffectiveTimeFactor);
udiChuckCloseTime := TIME_TO_UDINT(tChuckCloseTime) / TO_UDINT(uiEffectiveTimeFactor);
udiCycleStartTime := UDINT#200 / TO_UDINT(uiEffectiveTimeFactor);
udiCycleTime := TIME_TO_UDINT(tCycleTime) / TO_UDINT(uiEffectiveTimeFactor);

IF udiDoorOpenTime < UDINT#1 THEN udiDoorOpenTime := UDINT#1; END_IF;
IF udiDoorCloseTime < UDINT#1 THEN udiDoorCloseTime := UDINT#1; END_IF;
IF udiChuckOpenTime < UDINT#1 THEN udiChuckOpenTime := UDINT#1; END_IF;
IF udiChuckCloseTime < UDINT#1 THEN udiChuckCloseTime := UDINT#1; END_IF;
IF udiCycleStartTime < UDINT#1 THEN udiCycleStartTime := UDINT#1; END_IF;
IF udiCycleTime < UDINT#1 THEN udiCycleTime := UDINT#1; END_IF;

tEffectiveDoorOpenTime := UDINT_TO_TIME(udiDoorOpenTime);
tEffectiveDoorCloseTime := UDINT_TO_TIME(udiDoorCloseTime);
tEffectiveChuckOpenTime := UDINT_TO_TIME(udiChuckOpenTime);
tEffectiveChuckCloseTime := UDINT_TO_TIME(udiChuckCloseTime);
tEffectiveCycleStartTime := UDINT_TO_TIME(udiCycleStartTime);
tEffectiveCycleTime := UDINT_TO_TIME(udiCycleTime);

// =====================================================
// Первичная инициализация
// =====================================================

IF NOT xInitialized THEN
    Status.xDoorOpen := FALSE;
    Status.xDoorClosed := TRUE;
	Status.xHatchLocked := TRUE;
	Status.xSafetyDoorOpen := FALSE;
	Status.xSafetyDoorClosed := TRUE;

    Status.xChuckClamped := TRUE;
    Status.xChuckUnclamped := FALSE;

    Status.xCycleActive := FALSE;
    Status.xCycleDone := FALSE;
    Status.xAlarm := FALSE;

    xInitialized := TRUE;
END_IF;

IF xTestInitialize THEN
	xDoorOpening := FALSE;
	xDoorClosing := FALSE;
	xHatchUnlocking := FALSE;
	xSafetyDoorOpening := FALSE;
	xSafetyDoorClosing := FALSE;
	xChuckClamping := FALSE;
	xChuckOpening := FALSE;
	xCycleStarting := FALSE;
	xAlarmLatched := FALSE;
	Status.xDoorOpen := FALSE;
	Status.xDoorClosed := TRUE;
	Status.xHatchLocked := TRUE;
	Status.xSafetyDoorOpen := FALSE;
	Status.xSafetyDoorClosed := TRUE;
	Status.xChuckClamped := (uiTestInitialState = UINT#2) OR (uiTestInitialState = UINT#3);
	Status.xChuckUnclamped := NOT Status.xChuckClamped;
	Status.xCycleActive := uiTestInitialState = UINT#2;
	Status.xCycleDone := uiTestInitialState = UINT#3;
	Status.xAlarm := FALSE;
	Error.dwErrorActive := DWORD#0;
END_IF;

// Инъекция имеет приоритет над ручной командой закрытия. После снятия инъекции
// дверь остаётся открыта, пока оператор явно не подаст команду закрытия.
IF xSafetyDoorOpen THEN
	Status.xSafetyDoorOpen := TRUE;
	Status.xSafetyDoorClosed := FALSE;
	xSafetyDoorOpening := FALSE;
	xSafetyDoorClosing := FALSE;
END_IF;


// =====================================================
// Детектор запуска цикла
// =====================================================

rtStartCycle(CLK := Command.xStartCycle);


// =====================================================
// Формирование и сброс аварии
// =====================================================

xResetRequest := FaultRequest.xReset OR Command.xReset;

IF FaultRequest.xEnabled AND FaultRequest.xMachineAlarm THEN
	Error.dwErrorActive := Error.dwErrorActive OR ERR_MACHINE_ALARM;
END_IF;

IF FaultRequest.xEnabled
AND FaultRequest.xDoorFault
AND (xDoorOpening OR xDoorClosing) THEN
	Error.dwErrorActive := Error.dwErrorActive OR ERR_DOOR_FAULT;
END_IF;

IF FaultRequest.xEnabled
AND FaultRequest.xChuckFault
AND (xChuckClamping OR xChuckOpening) THEN
	Error.dwErrorActive := Error.dwErrorActive OR ERR_CHUCK_FAULT;
END_IF;

IF xResetRequest
AND NOT (FaultRequest.xEnabled AND FaultRequest.xMachineAlarm)
AND NOT (FaultRequest.xEnabled AND FaultRequest.xDoorFault)
AND NOT (FaultRequest.xEnabled AND FaultRequest.xChuckFault) THEN
	Error.dwErrorLast := Error.dwErrorActive;
	Error.dwErrorActive := DWORD#0;
END_IF;

// Отдельный сброс симулятора также отменяет зависшее тестовое действие.
// Штатный Command.xReset сохраняет прежнее поведение и только снимает ошибку.
IF FaultRequest.xReset THEN
	xDoorOpening := FALSE;
	xDoorClosing := FALSE;
	xHatchUnlocking := FALSE;
	xSafetyDoorOpening := FALSE;
	xSafetyDoorClosing := FALSE;
	xChuckClamping := FALSE;
	xChuckOpening := FALSE;
	xCycleStarting := FALSE;
END_IF;

xAlarmLatched := Error.dwErrorActive <> DWORD#0;


// =====================================================
// Приём команд станка
// =====================================================

IF NOT xAlarmLatched THEN

	// xHatchUnLock — единственный выход замка: TRUE снимает замок,
	// FALSE после закрытия двери возвращает его в безопасное состояние.
	IF Command.xHatchUnLock
	AND Status.xHatchLocked
	AND NOT Status.xCycleActive THEN
		xHatchUnlocking := TRUE;
	END_IF;
	IF NOT Command.xHatchUnLock
	AND Status.xDoorClosed THEN
		xHatchUnlocking := FALSE;
		Status.xHatchLocked := TRUE;
	END_IF;

    // Открытие двери
    IF Command.xOpenDoor
    AND NOT Status.xDoorOpen
    AND NOT Status.xCycleActive THEN
        xDoorOpening := TRUE;
        xDoorClosing := FALSE;
    END_IF;

    // Закрытие двери
    IF Command.xCloseDoor
    AND NOT Status.xDoorClosed THEN
        xDoorClosing := TRUE;
        xDoorOpening := FALSE;
    END_IF;

	// Операторская дверь не участвует в автоматическом рецепте и двигается
	// только отдельными ручными командами.
	IF Command.xOpenSafetyDoor
	AND NOT Status.xSafetyDoorOpen
	AND NOT Status.xCycleActive THEN
		xSafetyDoorOpening := TRUE;
		xSafetyDoorClosing := FALSE;
	END_IF;

	IF Command.xCloseSafetyDoor
	AND NOT Status.xSafetyDoorClosed
	AND NOT xSafetyDoorOpen
	AND NOT Status.xCycleActive THEN
		xSafetyDoorClosing := TRUE;
		xSafetyDoorOpening := FALSE;
	END_IF;

    // Зажим патрона
    IF Command.xClampChuck
    AND NOT Status.xChuckClamped
    AND NOT Status.xCycleActive THEN
        xChuckClamping := TRUE;
        xChuckOpening := FALSE;
    END_IF;

    // Разжим патрона
    IF Command.xUnclampChuck
    AND NOT Status.xChuckUnclamped
    AND NOT Status.xCycleActive THEN
        xChuckOpening := TRUE;
        xChuckClamping := FALSE;
    END_IF;

    // Запуск обработки
    IF rtStartCycle.Q
    AND Status.xDoorClosed
    AND Status.xChuckClamped
    AND NOT Status.xCycleActive THEN
        xCycleStarting := TRUE;
        Status.xCycleDone := FALSE;
    END_IF;

END_IF;


// =====================================================
// Таймеры механизмов
// =====================================================

tonDoorOpen(
    IN := xDoorOpening
		AND NOT (FaultRequest.xEnabled AND FaultRequest.xDoorFault),
	PT := tEffectiveDoorOpenTime
);

tonDoorClose(
    IN := xDoorClosing
		AND NOT (FaultRequest.xEnabled AND FaultRequest.xDoorFault),
	PT := tEffectiveDoorCloseTime
);

tonHatchUnlock(
	IN := xHatchUnlocking
		AND NOT (FaultRequest.xEnabled AND FaultRequest.xTimeoutHatchUnlock),
	PT := T#200MS
);

tonSafetyDoorOpen(
	IN := xSafetyDoorOpening,
	PT := tEffectiveDoorOpenTime
);

tonSafetyDoorClose(
	IN := xSafetyDoorClosing AND NOT xSafetyDoorOpen,
	PT := tEffectiveDoorCloseTime
);

tonChuckClamp(
    IN := xChuckClamping
		AND NOT (FaultRequest.xEnabled AND FaultRequest.xChuckFault),
	PT := tEffectiveChuckCloseTime
);

tonChuckOpen(
    IN := xChuckOpening
		AND NOT (FaultRequest.xEnabled AND FaultRequest.xChuckFault),
	PT := tEffectiveChuckOpenTime
);

tonCycleStart(
    IN := xCycleStarting,
    PT := tEffectiveCycleStartTime
);

tonCycle(
    IN := Status.xCycleActive AND NOT xAlarmLatched,
    PT := tEffectiveCycleTime
);


// =====================================================
// Завершение открытия двери
// =====================================================

IF tonDoorOpen.Q THEN
    Status.xDoorOpen := TRUE;
    Status.xDoorClosed := FALSE;

    xDoorOpening := FALSE;
END_IF;


// =====================================================
// Завершение закрытия двери
// =====================================================

IF tonDoorClose.Q THEN
    Status.xDoorClosed := TRUE;
    Status.xDoorOpen := FALSE;

    xDoorClosing := FALSE;
END_IF;

IF tonHatchUnlock.Q THEN
	Status.xHatchLocked := FALSE;
	xHatchUnlocking := FALSE;
END_IF;

// =====================================================
// Завершение движения операторской двери
// =====================================================

IF tonSafetyDoorOpen.Q THEN
	Status.xSafetyDoorOpen := TRUE;
	Status.xSafetyDoorClosed := FALSE;
	xSafetyDoorOpening := FALSE;
END_IF;

IF tonSafetyDoorClose.Q THEN
	Status.xSafetyDoorClosed := TRUE;
	Status.xSafetyDoorOpen := FALSE;
	xSafetyDoorClosing := FALSE;
END_IF;


// =====================================================
// Завершение зажима патрона
// =====================================================

IF tonChuckClamp.Q THEN
    Status.xChuckClamped := TRUE;
    Status.xChuckUnclamped := FALSE;

    xChuckClamping := FALSE;
END_IF;


// =====================================================
// Завершение разжима патрона
// =====================================================

IF tonChuckOpen.Q THEN
    Status.xChuckUnclamped := TRUE;
    Status.xChuckClamped := FALSE;

    xChuckOpening := FALSE;
END_IF;


// =====================================================
// Запуск цикла
// =====================================================

IF tonCycleStart.Q THEN
    Status.xCycleActive := TRUE;
    xCycleStarting := FALSE;
END_IF;


// =====================================================
// Завершение цикла
// =====================================================

IF tonCycle.Q THEN
    Status.xCycleActive := FALSE;
    Status.xCycleDone := TRUE;
END_IF;


// =====================================================
// Реакция на аварийное состояние
// =====================================================

IF xAlarmLatched THEN
    Status.xCycleActive := FALSE;

    xDoorOpening := FALSE;
    xDoorClosing := FALSE;
	xHatchUnlocking := FALSE;
	xSafetyDoorOpening := FALSE;
	xSafetyDoorClosing := FALSE;

    xChuckClamping := FALSE;
    xChuckOpening := FALSE;

    xCycleStarting := FALSE;
END_IF;


// =====================================================
// Выходной статус
// =====================================================

Status.xAlarm := xAlarmLatched;
Status.xReady := NOT xAlarmLatched
	AND NOT Status.xCycleActive
	AND NOT xDoorOpening
	AND NOT xDoorClosing
	AND NOT xHatchUnlocking
	AND NOT xSafetyDoorOpening
	AND NOT xSafetyDoorClosing
	AND NOT xChuckClamping
	AND NOT xChuckOpening;

Diag.xDoorOpening := xDoorOpening;
Diag.xDoorClosing := xDoorClosing;
Diag.xSafetyDoorOpening := xSafetyDoorOpening;
Diag.xSafetyDoorClosing := xSafetyDoorClosing;
Diag.xChuckClamping := xChuckClamping;
Diag.xChuckOpening := xChuckOpening;
Diag.xCycleStarting := xCycleStarting;
Diag.xResetAllowed := (Error.dwErrorActive <> DWORD#0)
	AND NOT (FaultRequest.xEnabled AND FaultRequest.xMachineAlarm)
	AND NOT (FaultRequest.xEnabled AND FaultRequest.xDoorFault)
	AND NOT (FaultRequest.xEnabled AND FaultRequest.xChuckFault);

IF Error.dwErrorActive <> DWORD#0 THEN
	Error.dwErrorLast := Error.dwErrorActive;
END_IF;

Error.stErrorActive := UpdateErrorView(dwError := Error.dwErrorActive);
Error.stErrorLast := UpdateErrorView(dwError := Error.dwErrorLast);

METHOD UpdateErrorView : ST_MACHINE_SIM_ERROR
VAR_INPUT
	dwError : DWORD; // Битовая маска для расшифровки
END_VAR
VAR
	stError : ST_MACHINE_SIM_ERROR; // Представление ошибок отдельными флагами
END_VAR
stError.MACHINE_ALARM := (dwError AND ERR_MACHINE_ALARM) <> DWORD#0;
stError.DOOR_FAULT := (dwError AND ERR_DOOR_FAULT) <> DWORD#0;
stError.CHUCK_FAULT := (dwError AND ERR_CHUCK_FAULT) <> DWORD#0;

UpdateErrorView := stError;
END_METHOD

END_FUNCTION_BLOCK

// Device/Application/FB/FB_FAULT_INJECTOR/FB_MACHINE_FAULT_INJECTOR
FUNCTION_BLOCK FB_MACHINE_FAULT_INJECTOR
VAR_INPUT
	Request            : ST_MACHINE_FAULT_REQUEST; // Запросы диагностической инъекции
	MachineStatusRaw    : ST_MACHINE_IO_STATUS; // Неизменённая обратная связь станка
	RobotStatusRaw      : ST_ROBOT_STATUS; // Неизменённая обратная связь робота
	NominalTimeouts     : ST_MACHINE_TIMEOUTS; // Штатные таймауты автомата станка
END_VAR
VAR_OUTPUT
	MachineStatus : ST_MACHINE_IO_STATUS; // Обратная связь, передаваемая FB_MACHINE
	RobotStatus   : ST_ROBOT_STATUS; // Статус робота, передаваемый FB_MACHINE
	Timeouts      : ST_MACHINE_TIMEOUTS; // Действующий профиль таймаутов
	Status        : ST_FAULT_INJECTION_STATUS; // Состояние источника для HMI
END_VAR
VAR CONSTANT
	SIMULATION_TIMEOUT : TIME := T#2S; // Ускоренное время диагностического сценария
END_VAR

// Инжектор не формирует маски ошибок. Он только искажает подтверждения,
// после чего FB_MACHINE обнаруживает штатный TIMEOUT собственными таймерами.

MachineStatus := MachineStatusRaw;
RobotStatus := RobotStatusRaw;
Timeouts := NominalTimeouts;

// Состояние источника аварии не должно оставаться активным после снятия
// соответствующего переключателя. Сам FB_MACHINE при этом сохраняет свою
// защёлкнутую ошибку и сбрасывается отдельной командой из меню станка.
MachineStatus.xAlarm := MachineStatusRaw.xAlarm
	AND Request.xEnabled
	AND (Request.xMachineAlarm OR Request.xDoorFault OR Request.xChuckFault);

Status.xAllowed := Request.xEnabled;
Status.xActive := Request.xEnabled AND (
	Request.xMachineAlarm
	OR Request.xDoorFault
	OR Request.xChuckFault
	OR Request.xTimeoutRobotMove
	OR Request.xTimeoutRobotAction
	OR Request.xTimeoutRobotRelease
	OR Request.xTimeoutDoorOpen
		OR Request.xTimeoutDoorClose
		OR Request.xTimeoutHatchUnlock
	OR Request.xTimeoutChuckOpen
	OR Request.xTimeoutChuckClose
	OR Request.xTimeoutCycleStart
);
Status.xBusy := FALSE;
Status.xResetAllowed := FALSE;
Status.xRejected := FALSE;

IF Request.xEnabled THEN
	IF Request.xTimeoutRobotMove THEN
		RobotStatus.xDone := FALSE;
		Timeouts.tRobotMove := SIMULATION_TIMEOUT;
	END_IF;

	IF Request.xTimeoutRobotAction THEN
		RobotStatus.xDone := FALSE;
		RobotStatus.xGripper1Open := FALSE;
		RobotStatus.xGripper1Closed := FALSE;
		RobotStatus.xGripper2Open := FALSE;
		RobotStatus.xGripper2Closed := FALSE;
		RobotStatus.xRotatedToBlank := FALSE;
		RobotStatus.xRotatedToDetail := FALSE;
		Timeouts.tRobotAction := SIMULATION_TIMEOUT;
	END_IF;

	IF Request.xTimeoutRobotRelease THEN
		RobotStatus.xBusy := TRUE;
		Timeouts.tRobotRelease := SIMULATION_TIMEOUT;
	END_IF;

	IF Request.xTimeoutDoorOpen THEN
		MachineStatus.xDoorOpen := FALSE;
		Timeouts.tDoorOpen := SIMULATION_TIMEOUT;
	END_IF;

	IF Request.xTimeoutDoorClose THEN
		MachineStatus.xDoorClosed := FALSE;
		Timeouts.tDoorClose := SIMULATION_TIMEOUT;
	END_IF;

	IF Request.xTimeoutHatchUnlock THEN
		MachineStatus.xHatchLocked := TRUE;
		Timeouts.tHatchUnlock := SIMULATION_TIMEOUT;
	END_IF;

	IF Request.xTimeoutChuckOpen THEN
		MachineStatus.xChuckUnclamped := FALSE;
		Timeouts.tChuckOpen := SIMULATION_TIMEOUT;
	END_IF;

	IF Request.xTimeoutChuckClose THEN
		MachineStatus.xChuckClamped := FALSE;
		Timeouts.tChuckClose := SIMULATION_TIMEOUT;
	END_IF;

	IF Request.xTimeoutCycleStart THEN
		MachineStatus.xCycleActive := FALSE;
		Timeouts.tCycleStart := SIMULATION_TIMEOUT;
	END_IF;
END_IF;

END_FUNCTION_BLOCK

// Device/Application/FB/FB_TWO_PALLET
FUNCTION_BLOCK FB_TWO_PALLET
VAR_INPUT
	xSelected : BOOL;
	xManual : BOOL;
	xSafe : BOOL;
	xRobotSwapWindow : BOOL; // Робот не выполняет и не ожидает операцию именно с этим магазином
	xRobotOperation : BOOL; // Текущая или уже выданная операция с этим магазином
	xPointsConfigured : BOOL; // Собственная база магазина нужна для ввода в автомат
	xRobotGeometryReady : BOOL; // Собственная база магазина и поддерживаемый интерфейс робота
	xRobotMagazineReady : BOOL; // Ошибки и геометрия магазина; содержимое не блокирует включение
	xConnection : BOOL; // Heartbeat HMI нужен только для ручных команд
	xStopRequest : BOOL; // Общий Stop прерывает движение, но не отключает неподвижный магазин
	xAutoSwap : BOOL;
	xOtherLoaded : BOOL;
	xActivePalletEditAllowed : BOOL;
	xConfigurationChanged : BOOL;
    xIoPneumaticOverride : BOOL; // Прямое воздействие на катушки снимает подтверждение расстановки
	xExternalCommandRejected : BOOL;
	Command : ST_TWO_PALLET_COMMAND;
	Config : ST_TWO_PALLET_CONFIG;
	Input : ST_TWO_PALLET_INPUT;
END_VAR
VAR_OUTPUT
	Status : ST_TWO_PALLET_STATUS;
	Diag : ST_TWO_PALLET_DIAG;
	Error : ST_TWO_PALLET_ERRORS;
	Output : ST_TWO_PALLET_OUTPUT;
END_VAR
VAR
	ePreviousState : E_TWO_PALLET_STATE := E_TWO_PALLET_STATE.IDLE;
	uiFrom : UINT;
	uiTo : UINT;
	uiSelected : UINT;
	uiCandidate : UINT;
	uiPreviousCandidate : UINT;
	uiConfirmedCandidate : UINT;
	uiManualSelected : UINT;
	uiJogDirection : UINT;
	uiSignals : UINT;
	uiSelectedSignals : UINT;
	uiTargetSignals : UINT;
	xPreviousBaseValid : BOOL;
	xConfigValid : BOOL;
	xContradiction : BOOL;
	xPairValid : BOOL;
	xWork : BOOL;
	xExchange : BOOL;
	xIdle : BOOL;
	xBase : BOOL;
	xRecovery : BOOL;
	xPneumaticBase : BOOL;
	xPneumaticRecovery : BOOL;
	xManualPneumaticState : BOOL;
	xAutomaticState : BOOL;
	xAxisMotionState : BOOL;
	xManualState : BOOL;
	xEnableBaseAllowed : BOOL;
	xAutoSwapAllowed : BOOL;
	xExchangeStartedManual : BOOL; // Обмен начат в ручном режиме: без проверки роботной зоны/точек
	xCommandPresent : BOOL;
	xAccepted : BOOL;
	xStateEntry : BOOL;
	xSeenMotion : BOOL;
	xSeenDone : BOOL;
	xLiftUpCommand : BOOL;
	xLiftDownCommand : BOOL;
	xSelectCommand : BOOL;
	xManualLockCommand : BOOL;
	xManualStopCommand : BOOL;
	xManualLockOutTarget : BOOL;
	xManualStopOutTarget : BOOL;
	xLockOutTarget : BOOL;
	xStopOutTarget : BOOL;
	xStartupInitialized : BOOL;
	xTrustedAtScanStart : BOOL;
	lrWork : LREAL;
	lrTarget : LREAL;
	lrSpan : LREAL;
	rTravel : REAL;
	tStateLimit : TIME;
	tonState : TON;
	tonCoil : TON;
	tonJogLease : TON;
	dwPreviousError : DWORD;
END_VAR
VAR CONSTANT
	ERR_DRIVE : DWORD := DWORD#16#100;
	ERR_SENSOR_CONTRADICTION : DWORD := DWORD#16#200;
	ERR_CYLINDER_TIMEOUT : DWORD := DWORD#16#400;
	ERR_MOTION_TIMEOUT : DWORD := DWORD#16#800;
	ERR_LOGIC : DWORD := DWORD#16#1000;
	ERR_SEQUENCE_INTERRUPTED : DWORD := DWORD#16#2000;
	WRN_COMMAND_REJECTED : UINT := UINT#30;
	WRN_ENABLE_POINTS : UINT := UINT#18; // Общий код с FB_MAGAZINE для отсутствующей базы
	WRN_START_REJECTED_BY_OPERATOR : UINT := UINT#31;
	JOG_POSITIVE : UINT := UINT#1;
	JOG_NEGATIVE : UINT := UINT#2;
END_VAR

// Шаги, разрешения и подтверждение положения не восстанавливаются после старта PLC.
IF NOT xStartupInitialized THEN
	Diag.eState := E_TWO_PALLET_STATE.IDLE;
	ePreviousState := E_TWO_PALLET_STATE.IDLE;
	Status.xConfirmed := FALSE;
	Status.xEnabled := FALSE;
	xStartupInitialized := TRUE;
END_IF;

Status.xCompleted := FALSE;
Status.Input := Input;
xTrustedAtScanStart := Status.xConfirmed;

// Все выходные команды импульсные или формируются заново на каждом скане.
Output.xPowerOn := FALSE;
Output.xPowerOff := FALSE;
Output.xDriveReset := FALSE;
Output.xHome := FALSE;
Output.xMove := FALSE;
Output.xStop := FALSE;
Output.xJogPositive := FALSE;
Output.xJogNegative := FALSE;
Output.xTeachOperator := FALSE;
Output.xTeachWork := FALSE;
xLiftUpCommand := FALSE;
xLiftDownCommand := FALSE;
xSelectCommand := FALSE;
xManualLockCommand := FALSE;
xManualStopCommand := FALSE;

// Конфигурация механизма.
xConfigValid := Config.xConfigured
	AND Config.xSignalPatternsConfigured
	AND IsSignalConfigurationValid(uiP1Signals := Config.uiP1Signals, uiP2Signals := Config.uiP2Signals)
	AND (Config.lrTolerance > 0.0)
	AND (Config.lrTolerance <= 20.0)
	AND (ABS(Config.lrWorkP1 - Config.lrExchange) > 2.0 * Config.lrTolerance)
	AND (ABS(Config.lrWorkP2 - Config.lrExchange) > 2.0 * Config.lrTolerance)
	AND ((Config.lrWorkP1 - Config.lrExchange) * (Config.lrWorkP2 - Config.lrExchange) > 0.0)
	AND (Config.lrVelocity > 0.0)
	AND (Config.lrAcceleration > 0.0)
	AND (Config.lrDeceleration > 0.0)
	AND (Config.lrJerk > 0.0)
	AND (Config.tPulse >= T#50MS)
	AND (Config.tCylinder > Config.tPulse)
	AND (Config.tMove > T#0S)
	AND (Config.tHome > T#0S);
Status.xConfigValid := xConfigValid;

// Фактическое состояние пневматики и каретки.
xContradiction := (Input.xLiftUp AND Input.xLiftDown)
	OR (Input.xLockIn AND Input.xLockOut)
	OR (Input.xStopIn AND Input.xStopOut)
	OR (Input.xLimitNegative AND Input.xLimitPositive);
xPairValid := (Input.xLockIn XOR Input.xLockOut)
	AND (Input.xStopIn XOR Input.xStopOut);

uiSignals := UINT#0;
IF Input.xLiftDown THEN uiSignals := uiSignals OR UINT#1; END_IF;
IF Input.xLiftUp THEN uiSignals := uiSignals OR UINT#2; END_IF;
IF Input.xLockIn THEN uiSignals := uiSignals OR UINT#4; END_IF;
IF Input.xLockOut THEN uiSignals := uiSignals OR UINT#8; END_IF;
IF Input.xStopIn THEN uiSignals := uiSignals OR UINT#16; END_IF;
IF Input.xStopOut THEN uiSignals := uiSignals OR UINT#32; END_IF;

uiSelected := UINT#0;
IF xPairValid THEN
	IF (uiSignals AND UINT#60) = (Config.uiP1Signals AND UINT#60) THEN
		uiSelected := UINT#1;
	ELSIF (uiSignals AND UINT#60) = (Config.uiP2Signals AND UINT#60) THEN
		uiSelected := UINT#2;
	END_IF;
END_IF;
xPairValid := xPairValid AND (uiSelected <> UINT#0);

lrWork := Config.lrWorkP1;
uiSelectedSignals := Config.uiP1Signals;
IF uiSelected = UINT#2 THEN
	lrWork := Config.lrWorkP2;
	uiSelectedSignals := Config.uiP2Signals;
END_IF;

xWork := xConfigValid
	AND Input.xHomed
	AND Input.xStandstill
	AND xPairValid
	AND (ABS(Input.lrPosition - lrWork) <= Config.lrTolerance);
xExchange := xConfigValid
	AND Input.xHomed
	AND Input.xStandstill
	AND (ABS(Input.lrPosition - Config.lrExchange) <= Config.lrTolerance);

uiCandidate := UINT#0;
IF xWork
	AND (uiSignals = uiSelectedSignals)
	AND NOT xContradiction
	AND NOT Input.xDriveError
	AND NOT Status.xHomeRequired THEN
	uiCandidate := uiSelected;
END_IF;

xIdle := Diag.eState = E_TWO_PALLET_STATE.IDLE;
xAutomaticState := (Diag.eState = E_TWO_PALLET_STATE.AUTO_LOWER)
	OR (Diag.eState = E_TWO_PALLET_STATE.AUTO_MOVE_TO_EXCHANGE)
	OR (Diag.eState = E_TWO_PALLET_STATE.AUTO_SELECT_PALLET)
	OR (Diag.eState = E_TWO_PALLET_STATE.AUTO_MOVE_TO_WORK)
	OR (Diag.eState = E_TWO_PALLET_STATE.AUTO_RAISE);
xAxisMotionState := (Diag.eState = E_TWO_PALLET_STATE.AUTO_MOVE_TO_EXCHANGE)
	OR (Diag.eState = E_TWO_PALLET_STATE.AUTO_MOVE_TO_WORK)
	OR (Diag.eState = E_TWO_PALLET_STATE.MANUAL_MOVE)
	OR (Diag.eState = E_TWO_PALLET_STATE.MANUAL_HOME)
	OR (Diag.eState = E_TWO_PALLET_STATE.MANUAL_JOG);
xManualState := (Diag.eState = E_TWO_PALLET_STATE.MANUAL_LOWER)
	OR (Diag.eState = E_TWO_PALLET_STATE.MANUAL_RAISE)
	OR (Diag.eState = E_TWO_PALLET_STATE.MANUAL_SELECT_PALLET)
	OR (Diag.eState = E_TWO_PALLET_STATE.MANUAL_MOVE)
	OR (Diag.eState = E_TWO_PALLET_STATE.MANUAL_HOME)
	OR (Diag.eState = E_TWO_PALLET_STATE.MANUAL_JOG)
	OR (Diag.eState = E_TWO_PALLET_STATE.MANUAL_LOCK)
	OR (Diag.eState = E_TWO_PALLET_STATE.MANUAL_STOP);
xManualPneumaticState := (Diag.eState = E_TWO_PALLET_STATE.MANUAL_LOWER)
	OR (Diag.eState = E_TWO_PALLET_STATE.MANUAL_LOCK)
	OR (Diag.eState = E_TWO_PALLET_STATE.MANUAL_STOP);

xBase := xSelected
	AND xConfigValid
	AND Input.xIoMapped
	AND Input.xAxisBound
	AND xSafe
	AND NOT xRobotOperation;
xRecovery := xBase
	AND xManual
	AND xConnection
	AND xIdle
	AND Input.xStandstill;
xPneumaticBase := xSelected
	AND xManual
	AND xSafe
	AND NOT xRobotOperation
	AND Input.xIoMapped
	AND Input.xStandstill;
xPneumaticRecovery := xPneumaticBase AND xIdle;

Status.uiCandidate := uiCandidate;
Status.uiSelected := uiSelected;

// Любое изменение достоверной расстановки аннулирует старое подтверждение.
IF (uiCandidate <> uiPreviousCandidate) OR (xBase <> xPreviousBaseValid) THEN
	Status.udiRevision := Status.udiRevision + UDINT#1;
	IF Status.udiRevision = UDINT#0 THEN
		Status.udiRevision := UDINT#1;
	END_IF;
END_IF;
uiPreviousCandidate := uiCandidate;
xPreviousBaseValid := xBase;

IF xConfigurationChanged THEN
	Status.xConfirmed := FALSE;
	Status.xEnabled := FALSE;
	Status.udiRevision := Status.udiRevision + UDINT#1;
	IF Status.udiRevision = UDINT#0 THEN
		Status.udiRevision := UDINT#1;
	END_IF;
END_IF;

IF xIoPneumaticOverride THEN
    Status.xConfirmed := FALSE;
    Status.xEnabled := FALSE;
    Status.udiRevision := Status.udiRevision + UDINT#1;
    IF Status.udiRevision = UDINT#0 THEN Status.udiRevision := UDINT#1; END_IF;
END_IF;

IF NOT xSelected
	OR NOT xSafe
	OR NOT Input.xAxisBound
	OR NOT Input.xIoMapped
	OR NOT xConfigValid
	OR Input.xDriveError
	OR NOT Input.xPowered
	OR (xIdle AND (uiCandidate <> uiConfirmedCandidate)) THEN
	Status.xConfirmed := FALSE;
END_IF;
// Первая невыполненная предпосылка для HMI.
Diag.uiReason := UINT#0;
IF NOT xSelected THEN
	Diag.uiReason := UINT#1;
ELSIF NOT xConfigValid THEN
	Diag.uiReason := UINT#2;
ELSIF NOT Input.xAxisBound OR NOT Input.xIoMapped THEN
	Diag.uiReason := UINT#3;
ELSIF NOT xSafe THEN
	Diag.uiReason := UINT#4;
ELSIF NOT xConnection THEN
	Diag.uiReason := UINT#17;
ELSIF Input.xDriveError THEN
	Diag.uiReason := UINT#6;
ELSIF Error.dwErrorActive <> DWORD#0 THEN
	Diag.uiReason := UINT#19;
ELSIF NOT Input.xPowered THEN
	Diag.uiReason := UINT#18;
ELSIF xContradiction THEN
	Diag.uiReason := UINT#7;
ELSIF Status.xHomeRequired OR NOT Input.xHomed THEN
	Diag.uiReason := UINT#8;
ELSIF NOT xPairValid THEN
	Diag.uiReason := UINT#9;
ELSIF NOT Input.xStandstill THEN
	Diag.uiReason := UINT#10;
ELSIF NOT xWork THEN
	Diag.uiReason := UINT#11;
ELSIF uiSignals <> uiSelectedSignals THEN
	Diag.uiReason := UINT#12;
ELSIF NOT xIdle THEN
	Diag.uiReason := UINT#22;
ELSIF NOT xRobotMagazineReady THEN
	Diag.uiReason := UINT#16;
ELSIF NOT xPointsConfigured THEN
	Diag.uiReason := UINT#15;
ELSIF NOT Status.xConfirmed AND NOT xManual THEN
	Diag.uiReason := UINT#20;
ELSIF NOT Status.xConfirmed THEN
	Diag.uiReason := UINT#13;
END_IF;

// Аварии механизма: биты 8..13 зарезервированы в MAGAZINE_LOGIC_1/2.
IF xSelected AND Input.xDriveError THEN
	Error.dwErrorActive := Error.dwErrorActive OR ERR_DRIVE;
	Status.xHomeRequired := TRUE;
END_IF;

IF xSelected AND xContradiction THEN
	Error.dwErrorActive := Error.dwErrorActive OR ERR_SENSOR_CONTRADICTION;
END_IF;

IF xSelected
	AND NOT xIdle
	AND (((NOT xBase) AND NOT (xManualPneumaticState AND xPneumaticBase))
		OR ((NOT xConnection) AND xManualState AND NOT xManualPneumaticState) OR xStopRequest
		OR (xAutomaticState AND ((xExchangeStartedManual AND NOT xManual)
			OR NOT xRobotSwapWindow))) THEN
	Error.dwErrorActive := Error.dwErrorActive OR ERR_SEQUENCE_INTERRUPTED;
	Diag.eState := E_TWO_PALLET_STATE.IDLE;
	Output.xStop := TRUE;
END_IF;

IF xSelected AND (xTrustedAtScanStart OR xAutomaticState) THEN
	IF ((Diag.eState <> E_TWO_PALLET_STATE.AUTO_SELECT_PALLET) AND NOT xPairValid)
		OR (((Diag.eState = E_TWO_PALLET_STATE.AUTO_MOVE_TO_EXCHANGE)
			OR (Diag.eState = E_TWO_PALLET_STATE.AUTO_MOVE_TO_WORK))
			AND (NOT Input.xLiftDown OR Input.xLiftUp))
		OR (xIdle AND (uiCandidate = UINT#0)) THEN
		Error.dwErrorActive := Error.dwErrorActive OR ERR_LOGIC;
	END_IF;
END_IF;

IF xSelected
	AND xTrustedAtScanStart
	AND (NOT xSafe
		OR NOT Input.xAxisBound
		OR NOT Input.xIoMapped
		OR NOT Input.xPowered) THEN
	Error.dwErrorActive := Error.dwErrorActive OR ERR_SEQUENCE_INTERRUPTED;
END_IF;

IF xSelected
	AND ((xContradiction AND NOT xIdle AND NOT xManualPneumaticState)
		OR (Input.xDriveError AND xAxisMotionState)) THEN
	Diag.eState := E_TWO_PALLET_STATE.IDLE;
	Output.xStop := TRUE;
END_IF;

IF xSelected AND NOT Input.xPowered AND (xAutomaticState OR xAxisMotionState) THEN
	Error.dwErrorActive := Error.dwErrorActive OR ERR_SEQUENCE_INTERRUPTED;
	Status.xHomeRequired := TRUE;
	Diag.eState := E_TWO_PALLET_STATE.IDLE;
	Output.xStop := TRUE;
END_IF;

IF Error.dwErrorActive <> DWORD#0 THEN
	Status.xEnabled := FALSE;
	Status.xConfirmed := FALSE;
	IF xAutomaticState THEN
		Diag.eState := E_TWO_PALLET_STATE.IDLE;
		Output.xStop := TRUE;
	END_IF;
END_IF;

